      |     #log_info("gripper config:",to_str(GRIPPER_CONFIG_MAP[i]))
      |     if (GRIPPER_CONFIG_MAP[i].object == objectname):
      |         log_info("found gripper parameters [" + to_str(GRIPPER_CONFIG_MAP[i]) + "]")
      |         return GRIPPER_CONFIG_MAP[i]
      |     end
      |     i = i + 1
      | end
      | 
      | log_warning("no gripper parameters found for object type: " + to_str(objectname))
      | return create_gripper_config()
      | end
      | # Function to find a landmark by item
      | def find_landmark_by_id(lm_id):
      |     local i = 0
      |     while i < LANDMARK_MAP.length():
      |         if LANDMARK_MAP[i].lm_id == lm_id:
      |             log_info("found landmark with id(" + to_str(lm_id) + "): [" + to_str(LANDMARK_MAP[i].description) + "]")
      |             return LANDMARK_MAP[i]
      |         end
      |         i = i + 1
      |     end
      |     log_warning("landmark not found for lm_id [" + to_str(lm_id) + "]")
      |     return create_landmark()
      | end
      | # Function to find a landmark by item
      | def find_landmark_by_capture_pos(capture_pos):
      |     local i = 0
      |     while i < LANDMARK_MAP.length():
      |         if LANDMARK_MAP[i].capture_pos == capture_pos:
      |             log_info("found landmark by capture_pos [" + to_str(LANDMARK_MAP[i].description) + "]")
      |             return LANDMARK_MAP[i]
      |         end
      |         i = i + 1
      |     end
      |     log_warning("Landmark not found for capture_pos: [" + to_str(capture_pos) + "]")
      |     return create_landmark()
      | end
      | 
      | def update_landmark_by_capture_pos(capture_pos, lm_pos):
      |     local i = 0
      |     while i < LANDMARK_MAP.length():
      |         if LANDMARK_MAP[i].capture_pos == capture_pos:
      |             log_info("updated landmark from [" + to_str(LANDMARK_MAP[i].description) + "]")
      |             LANDMARK_MAP[i].actual_frame = lm_pos
      |             return True
      |         end
      |         i = i + 1
      |     end
      |     log_warning("Landmark not found for capture_pos: [" + to_str(capture_pos) + "]")
      |     return False
      | end
      | 
      | def update_landmark_by_id(lm_id,lm_pos):
      |     local i = 0
      |     while i < LANDMARK_MAP.length():
      |         if LANDMARK_MAP[i].lm_id == lm_id:
      |             log_info("updated landmark.actual_frame from [" + to_str(LANDMARK_MAP[i].description + "]"))
      |             LANDMARK_MAP[i].actual_frame = lm_pos
      |             return True
      |         end
      |         i = i + 1
      |     end
      |     log_warning("Landmark not found for lm_id " + to_str(lm_id))
      |     return False
      | end
      | 
      | def find_vision_config_by_frame(frame):
      |     local i = 0
      |     while i < VISION_CONFIG_MAP.length():
      |         if VISION_CONFIG_MAP[i].capture_pos == frame:
      |             log_info("Vision Config found: [" + to_str(VISION_CONFIG_MAP[i].description) + "]")
      |             return VISION_CONFIG_MAP[i]
      |         end
      |         i = i + 1
      |     end
      |     log_info("Vision Config not found for frame: " + to_str(frame))
      |     return create_vision_config()
      | end
      | 
      | def find_vision_config_by_itemid(id):
      |     local i = 0
      |     while i < VISION_CONFIG_MAP.length():
      |         if VISION_CONFIG_MAP[i].item_id == id:
      |             log_info("Vision Config found: [" + to_str(VISION_CONFIG_MAP[i].description) + "]")
      |             return VISION_CONFIG_MAP[i]
      |         end
      |         i = i + 1
      |     end
      |     log_info("Vision Config not found for item: " + to_str(id))
      |     return create_vision_config()
      | end
      | 
      | def find_inspect_config_by_itemid(id):
      |     local i = 0
      |     while i < INSPECT_CONFIG_MAP.length():
      |         if INSPECT_CONFIG_MAP[i].item_id == id:
      |             log_info("Inspect Config found: [" + to_str(INSPECT_CONFIG_MAP[i].description) + "]")
      |             return INSPECT_CONFIG_MAP[i]
      |         end
      |         i = i + 1
      |     end
      |     log_info("Inspect Config not found for item: " + to_str(id))
      |     return create_inspect_config()
      | end
    Script file /programs/04 Scripts/SCRIPT Device Robotiq Greifer v0.2.script
      | # ############ SCRIPT Device Robotiq Greifer ###############
      | # **********************************************************
      | # Customer          :   URG
      | # Product Name      :   uLabMobile
      | # **********************************************************
      | # Controller/Robot  :   UR5e
      | # Software          :   5.17
      | # Dependencies      :   Logs Script, Robotiq Gripper and Gripper Datastructure for args (Factory Script), URCAP Robotiq
      | # **********************************************************
      | # Author            :   D.Kreugel, P.Köhnke
      | # Copyright (c)     :   United Robotics Group Health and Food GmbH
      | #                       An der Riede 2
      | #                       28816 Stuhr
      | #                       Germany
      | # *********************************************************
      | # Description       :   Gripper Robotiq Device Interface for Robotiq E-Hand Gripper
      | # Version           :   0.2
      | # Created           :   18.07.2024
      | # Updated           :
      | # *********************************************************
      | # Modifications     :
      | #
      | # Date              :
      | # Name              :
      | # Reason            :
      | # *********************************************************
      | # TODO              :   documentation
      | 
      | # RobotiQ Gripper
      | ROBOTIQ_GRP_CLOSE = 0
      | ROBOTIQ_GRP_OPEN = 40
      | 
      | # #############FORCEMODE###############
      | ROBOTIQ_GRP_FORCE = struct(FULL=100, HALF=50, LOW=25, NONE=0)
      | 
      | # #############SPEED###################
      | ROBOTIQ_GRP_SPEED = struct(FAST=100, MEDIUM=50, SLOW=20)
      | 
      | # ############VALIDATION###############
      | ROBOTIQ_GRP_VALIDATION = struct(ON=1, OFF=0, SKIP=-1)
      | 
      | # struct(prepick=0, pick=0, place=0, force=0, speed=0, validation=0, object_type=0, description="default")
      | def gripper_robotiq_activate():
      |     return rq_activate_and_wait()
      | end
      | 
      | def gripper_robotiq_reset_and_activate():
      |     return rq_reset_and_activate()
      |     #return rq_reset()
      | end
      | 
      | def gripper_robotiq_is_activated():
      |     return rq_is_gripper_activated()
      | end
      | 
      | def gripper_robotiq_get_current_pos_mm():
      |     return rq_current_pos_mm()
      | end
      | # Function to check if the RobotiQ gripper has an object
      | def gripper_robotiq_has_object():
      |     result = rq_is_object_detected()
      |     if result == False:
      |         log_error("No object detected by the gripper")
      |     end
      |     return result
      | end
      | 
      | def gripper_robotiq_move_to_mm(mm):
      |     if(gripper_robotiq_is_activated() == False):
      |         gripper_robotiq_activate()
      |     end
      |     return rq_move_and_wait_mm(mm)
      | end
      | 
      | def gripper_robotiq_close():
      |     if(gripper_robotiq_is_activated() == False):
      |         gripper_robotiq_activate()
      |     end
      |     return rq_close_and_wait()
      | end
      | 
      | def gripper_robotiq_open():
      |     if(gripper_robotiq_is_activated() == False):
      |         gripper_robotiq_activate()
      |     end
      |     return rq_open_and_wait()
      | end
      | 
      | def gripper_robotiq_set_force(force):
      |     return rq_set_force_norm(force)
      | end
      | 
      | def gripper_robotiq_set_speed(velocity):
      |     return rq_set_speed_norm(velocity)
      | end
      | # Function to initialize the RobotiQ gripper
      | # args = struct(obj_type = object.obj_type, force = force, speed = speed, validation = validation, width = (prepick=2, pick=0, place=2))
      | def gripper_robotiq_init(args):
      |     log_info("args:"+to_str(args))
      |     gripper_robotiq_set_force(args.force)
      |     gripper_robotiq_set_speed(args.speed)
      |     if(gripper_robotiq_is_activated() == False):
      |         gripper_robotiq_activate()
      |     end
      |     log_info("Robotiq Gripper Initialized with arguments:" + to_str(args))
      |     return True
      | end
      | # Function to prepare the RobotiQ gripper for picking
      | # args = struct(obj_type = object.obj_type, force = force, speed = speed, validation = validation, width = (prepick=2, pick=0, place=2))
      | def gripper_robotiq_prepick(args):
      |     gripper_robotiq_init(args)
      | 
      |     if(args.width.prepick <= ROBOTIQ_GRP_CLOSE):
      |         rq_close_and_wait()
      |     elif(args.width.prepick >= ROBOTIQ_GRP_OPEN):
      |         rq_open_and_wait()
      |     else:
      |         rq_move_and_wait_mm(args.width.prepick)
      |     end
      | 
      |     log_info("Robotiq Gripper prepick with arguments:" + to_str(args))
      |     return True
      | end
      | 
      | # Function to place an object using the RobotiQ gripper
      | # args = struct(obj_type = object.obj_type, force = force, speed = speed, validation = validation, width = (prepick=2, pick=0, place=2))
      | def gripper_robotiq_place(args):
      |     gripper_robotiq_init(args)
      | 
      |     if(args.width.place <= ROBOTIQ_GRP_CLOSE):
      |         rq_close_and_wait()
      |     elif(args.width.place >= ROBOTIQ_GRP_OPEN):
      |         rq_open_and_wait()
      |     else:
      |         rq_move_and_wait_mm(args.width.place)
      |     end
      | 
      |     log_info("Gripper Place with arguments:"+ to_str(args))
      |     return True
      | end
      | 
      | # Function to pick an object using the RobotiQ gripper
      | # args = struct(obj_type = object.obj_type, force = force, speed = speed, validation = validation, width = (prepick=2, pick=0, place=2))
      | def gripper_robotiq_pick(args):
      |     gripper_robotiq_init(args)
      | 
      |     if(args.width.pick <= ROBOTIQ_GRP_CLOSE):
      |         rq_close_and_wait()
      |     elif(args.width.pick >= ROBOTIQ_GRP_OPEN):
      |         rq_open_and_wait()
      |     else:
      |         rq_move_and_wait_mm(args.width.pick)
      |     end
      | 
      |     log_info("Gripper Pick with arguments:" + to_str(args))
      | 
      |     if args.validation == ROBOTIQ_GRP_VALIDATION.ON:
      |         if gripper_robotiq_has_object() == False:
      |             log_error("Validation failed, no object detected")
      |             return False
      |         end
      |     end
      | 
      |     return True
      | end
      | 
      | 
      | # def gripper_robotiq_close_and_validate():
      | #     rq_close_and_wait()
      | #     if gripper_robotiq_has_object() == False:
      | #         log_error("Validation failed, no object detected")
      | #         return False
      | #     else:
      | #         return True
      | #     end
      | # end
    Script file /programs/04 Scripts/SCRIPT uLM Gripperconfig v0.6.script
      | ############# SCRIPT uLM Gripperconfig ###############
      | #*****************************************************
      | # Customer          :   URG
      | # Product Name      :   uLabMobile
      | #****************************************************
      | # Controller/Robot  :   UR5e
      | # Software          :   UR-Script
      | # Dependencies      :   physical Gripper and Datastructure from Factory for args -> Device Script and Implementations of the Functions
      | # How To            :   Assign all Functioncalls to the equivalent of the used Device Script
      | #****************************************************
      | # Author            :   D.Kreugel, P.Köhnke
      | # Copyright (c)     :   United Robotics Group Health and Food GmbH
      | #                       An der Riede 2
      | #                       28816 Stuhr
      | #                       Germany
      | #****************************************************
      | # Description       :   Defines all Gripperm related Parameters and Functions
      | # Version           :   0.6
      | # Created           :   18.07.2024
      | # Updated           :
      | #****************************************************
      | # Modifications     :   -> at the moment Gripperconfig linked to Robotiq Gripper Device Script
      | # Date              :   18.07.2017
      | # Name              :   D.Kreugel
      | # Reason            :   uLM Standard
      | #****************************************************
      | # TO DO             : Implement Activate and Reset Routine at the beginning or after an error depending on the state if an Object is gripped or not, documentation
      | 
      | 
      | 
      | # GRIPPER DEFINES
      | GRIPPER_CLOSE = ROBOTIQ_GRP_CLOSE
      | GRIPPER_OPEN = ROBOTIQ_GRP_OPEN
      | # #############FORCE###############
      | GRIPPER_FORCE = ROBOTIQ_GRP_FORCE
      | # #############SPEED###################
      | GRIPPER_SPEED = ROBOTIQ_GRP_SPEED
      | # ############VALIDATION###############
      | GRIPPER_VALIDATION = ROBOTIQ_GRP_VALIDATION
      | 
      | # takes force in %
      | def gripper_set_force(force):
      |     return gripper_robotiq_set_force(force)
      | end
      | 
      | # takes speed in %
      | def gripper_set_speed(velocity):
      |     return gripper_robotiq_set_speed(velocity)
      | end
      | 
      | def gripper_activate():
      |     return gripper_robotiq_activate()
      | end
      | 
      | def gripper_reset_and_activate():
      |     return gripper_robotiq_reset_and_activate()
      | end
      | 
      | def gripper_is_activated():
      |     return gripper_robotiq_is_activated()
      | end
      | 
      | def gripper_get_current_pos_mm():
      |     return gripper_robotiq_get_current_pos_mm()
      | end
      | 
      | def gripper_has_object():
      |     return gripper_robotiq_has_object()
      | end
      | 
      | def gripper_open():
      |     return gripper_robotiq_open()
      | end
      | 
      | def gripper_close():
      |     return gripper_robotiq_close()
      | end
      | 
      | def gripper_move_to_pos_mm(mm):
      |     return gripper_robotiq_move_to_mm(mm)
      | end
      | 
      | # args = struct(obj_type = object.obj_type, force = force, speed = speed, validation = validation, width = (prepick=2, pick=0, place=2))
      | def gripper_init(args):
      |     return gripper_robotiq_init(args)
      | end
      | 
      | # args = struct(obj_type = object.obj_type, force = force, speed = speed, validation = validation, width = (prepick=2, pick=0, place=2))
      | def gripper_prepick(args):
      |     return gripper_robotiq_prepick(args)
      | end
      | 
      | # args = struct(obj_type = object.obj_type, force = force, speed = speed, validation = validation, width = (prepick=2, pick=0, place=2))
      | def gripper_pick(args):
      |     return gripper_robotiq_pick(args)
      | end
      | 
      | # args = struct(obj_type = object.obj_type, force = force, speed = speed, validation = validation, width = (prepick=2, pick=0, place=2))
      | def gripper_place(args):
      |     return gripper_robotiq_place(args)
      | end
      | 
      | 
      | # def gripper_close_and_validate():
      | #     return gripper_robotiq_close_and_validate()
      | # end
    Script file /programs/04 Scripts/SCRIPT uLM Projectconfig 0.2.script
      | ############# SCRIPT uLM Projectconfig ###############
      | #*****************************************************
      | # Customer          :   URG
      | # Product Name      :   uLabMobile
      | #****************************************************
      | # Controller/Robot  :   UR5e
      | # Software          :   5.17
      | # Dependencies      :   Factory Script, Defines Script, relevant project knowledge about objects, patterns, items, commands, vision skills, landmarktypes and movements
      | # How To            :   Define Step by Step all Project Data by creating the objects and appending them to the assigned List, if you skip information
      | #                       the default value will be assigned -> give as many details as possible as the default values will not work in some cases
      | #****************************************************
      | # Author            :   D.Kreugel
      | # Copyright (c)     :   United Robotics Group Health and Food GmbH
      | #                       An der Riede 2
      | #                       28816 Stuhr
      | #                       Germany
      | #****************************************************
      | # Description       :   Project Related Configurations -> in the future will be configured by UGO
      | # Version           :   0.2
      | # Created           :   18.07.2024
      | # Updated           :
      | #****************************************************
      | # Modifications     :
      | # Date              :
      | # Name              :
      | # Reason            :
      | #****************************************************
      | # TO DO             :  Simplify Rack Assignment, create Enums for Choices that can be made and will be repeated in many projects, documentation
      | 
      | #
      | 
      | # Please Import DeviceScripts and Defines Script First as you may wanna use some of the Defined Variables here
      | 
      | # Define here the Objects that should be handled, add a new Object Type in the defines if necessary
      | # create_object(id=0, obj_name=0, height=0, width=0, color="default", material="default", description="default")
      | # struct(NONE=0, CC_SAMPLE=1, CC_RACK=2, COAG_SAMPLE=3, COAG_RACK=4, HEMA_SAMPLE=5, HEMA_RACK=6, INPUT_RACK=7, CF_RACK=8, ANY_SAMPLE=9, ANY_RACK=10)
      | #create_object(id=0, obj_name=0, height=0, width=0, obj_type = 0, description="default")
      | OBJECT_MAP.append(create_object(id=0, obj_name=Objects.NONE, obj_type=ObjectType.NONE, height=0, width=0, description="None Object"))
      | OBJECT_MAP.append(create_object(id=1, obj_name=Objects.CC_SAMPLE, obj_type=ObjectType.SAMPLE, height=108, width=15, description="BD Li-Heparin"))
      | OBJECT_MAP.append(create_object(id=2, obj_name=Objects.HEMA_SAMPLE, obj_type=ObjectType.SAMPLE, height=81, width=13, description="BD EDTA"))
      | OBJECT_MAP.append(create_object(id=3, obj_name=Objects.CC_SAMPLE, obj_type=ObjectType.SAMPLE, height=108, width=15, description="BD Li-Heparin"))
      | OBJECT_MAP.append(create_object(id=4, obj_name=Objects.HEMA_SAMPLE, obj_type=ObjectType.SAMPLE, height=81, width=13, description="Sarstedt EDTA"))
      | OBJECT_MAP.append(create_object(id=5, obj_name=Objects.CC_SAMPLE, obj_type=ObjectType.SAMPLE, height=110, width=15, description="Sarstedt Serum-Gel"))
      | OBJECT_MAP.append(create_object(id=6, obj_name=Objects.ANY_SAMPLE, obj_type=ObjectType.SAMPLE, height=110, width=15, description="Any Sample"))
      | OBJECT_MAP.append(create_object(id=7, obj_name=Objects.ANY_RACK, height=150, width=120, description="Any Rack"))
      | OBJECT_MAP.append(create_object(id=8, obj_name=Objects.CF_RACK, height=110, width=15, description="Centrifuge Rack"))
      | OBJECT_MAP.append(create_object(id=12, obj_name=Objects.COBAS_RACK, height=OBJECT_REFERENCE_HEIGHT, width=20, description="Cobas Rack"))
      | OBJECT_MAP.append(create_object(id=9, obj_name=Objects.TARA_SAMPLE, obj_type=ObjectType.SAMPLE, height=110, width=15, description="Tara Sample"))
      | OBJECT_MAP.append(create_object(id=10, obj_name=Objects.BUTTON, obj_type=ObjectType.BUTTON, height=0, width=0, description="Button"))
      | OBJECT_MAP.append(create_object(id=11, obj_name=Objects.XN550_DRAWER, height=OBJECT_REFERENCE_HEIGHT, width=25, description="XN550 Drawer"))
      | 
      | #create_sample(obj_id=0, diameter=0, color="", material="", description="")
      | SAMPLES = make_list(0,create_sample(),MAX_ITEM_OBJ)
      | SAMPLES.append(create_sample(obj_id=1, cap_diameter=17.4, raw_diameter=15.3, color="darkgreen", material="88", description="BD Li-Heparin -> decapped in Cobas"))
      | SAMPLES.append(create_sample(obj_id=1, cap_diameter=17.4, raw_diameter=15.3, color="darkgreen", material="80", description="BD Li-Heparin -> decapped in Cobas"))
      | SAMPLES.append(create_sample(obj_id=1, cap_diameter=17.4, raw_diameter=15.3, color="darkgreen", material="93", description="BD Li-Heparin -> decapped in archive"))
      | SAMPLES.append(create_sample(obj_id=2, cap_diameter=15.5, raw_diameter=12.3, color="violet", material="82", description="BD EDTA -> Sysmex ->Archive"))
      | SAMPLES.append(create_sample(obj_id=2, cap_diameter=15.5, raw_diameter=12.3, color="violet", material="91", description="BD EDTA ->Archive"))
      | SAMPLES.append(create_sample(obj_id=2, cap_diameter=15.5, raw_diameter=12.3, color="violet", material="96", description="BD EDTA ->Archive"))
      | SAMPLES.append(create_sample(obj_id=3, cap_diameter=17.4, raw_diameter=15.3, color="lightgreen", material="88", description="BD Li-Heparin -> decapped in Cobas"))
      | SAMPLES.append(create_sample(obj_id=3, cap_diameter=17.4, raw_diameter=15.3, color="lightgreen", material="93", description="BD Li-Heparin -> decapped in Archive"))
      | SAMPLES.append(create_sample(obj_id=3, cap_diameter=17.4, raw_diameter=15.3, color="lightgreen", material="97", description="BD Li-Heparin -> decapped in Archive"))
      | SAMPLES.append(create_sample(obj_id=4, cap_diameter=15.6, raw_diameter=12.3, color="red", material="82", description="BD EDTA -> Sysmex ->Archive"))
      | SAMPLES.append(create_sample(obj_id=4, cap_diameter=15.6, raw_diameter=12.3, color="red", material="91", description="BD EDTA -> Archive"))
      | SAMPLES.append(create_sample(obj_id=4, cap_diameter=15.6, raw_diameter=12.3, color="red", material="96", description="BD EDTA -> Archive"))
      | SAMPLES.append(create_sample(obj_id=5, cap_diameter=17.4, raw_diameter=15.3, color="brown", material="80", description="Sarstedt Serum-Gel -> decapped in Cobas"))
      | SAMPLES.append(create_sample(obj_id=5, cap_diameter=17.4, raw_diameter=15.3, color="brown", material="93", description="Sarstedt Serum-Gel -> decapped in Archive"))
      | 
      | # Gripper Configurations depending on the Object Type , add new force and speed in the Defines if necessary
      | # create_gripper_config(gripper_offset=struct(prepick=2, pick=0, place=2), force=0, speed=0, validation=0, object=create_object())
      | GRIPPER_CONFIG_MAP.append(create_gripper_config(gripper_offset=struct(prepick=2, pick=0, place=2), force=GRIPPER_FORCE.HALF, speed=GRIPPER_SPEED.MEDIUM, validation=GRIPPER_VALIDATION.ON, object=find_object_by_objectname(Objects.ANY_SAMPLE)))
      | GRIPPER_CONFIG_MAP.append(create_gripper_config(gripper_offset=struct(prepick=2, pick=0, place=2), force=GRIPPER_FORCE.FULL, speed=GRIPPER_SPEED.MEDIUM, validation=GRIPPER_VALIDATION.ON, object=find_object_by_objectname(Objects.ANY_RACK)))
      | GRIPPER_CONFIG_MAP.append(create_gripper_config(gripper_offset=struct(prepick=2, pick=0, place=2), force=GRIPPER_FORCE.HALF, speed=GRIPPER_SPEED.MEDIUM, validation=GRIPPER_VALIDATION.ON, object=find_object_by_objectname(Objects.CC_SAMPLE)))
      | GRIPPER_CONFIG_MAP.append(create_gripper_config(gripper_offset=struct(prepick=3, pick=0, place=3), force=GRIPPER_FORCE.HALF, speed=GRIPPER_SPEED.MEDIUM, validation=GRIPPER_VALIDATION.ON, object=find_object_by_objectname(Objects.HEMA_SAMPLE)))
      | GRIPPER_CONFIG_MAP.append(create_gripper_config(gripper_offset=struct(prepick=4, pick=0, place=4), force=GRIPPER_FORCE.HALF, speed=GRIPPER_SPEED.MEDIUM, validation=GRIPPER_VALIDATION.OFF, object=find_object_by_objectname(Objects.TARA_SAMPLE)))
      | GRIPPER_CONFIG_MAP.append(create_gripper_config(gripper_offset=struct(prepick=2, pick=0, place=2), force=GRIPPER_FORCE.FULL, speed=GRIPPER_SPEED.MEDIUM, validation=GRIPPER_VALIDATION.ON, object=find_object_by_objectname(Objects.CF_RACK)))
      | GRIPPER_CONFIG_MAP.append(create_gripper_config(gripper_offset=struct(prepick=2, pick=0, place=2), force=GRIPPER_FORCE.FULL, speed=GRIPPER_SPEED.MEDIUM, validation=GRIPPER_VALIDATION.ON, object=find_object_by_objectname(Objects.COBAS_RACK)))
      | GRIPPER_CONFIG_MAP.append(create_gripper_config(gripper_offset=struct(prepick=0, pick=0, place=0), force=GRIPPER_FORCE.HALF, speed=GRIPPER_SPEED.MEDIUM, validation=GRIPPER_VALIDATION.OFF, object=find_object_by_objectname(Objects.NONE)))
      | GRIPPER_CONFIG_MAP.append(create_gripper_config(gripper_offset=struct(prepick=0, pick=0, place=0), force=GRIPPER_FORCE.HALF, speed=GRIPPER_SPEED.MEDIUM, validation=GRIPPER_VALIDATION.OFF, object=find_object_by_objectname(Objects.BUTTON)))
      | GRIPPER_CONFIG_MAP.append(create_gripper_config(gripper_offset=struct(prepick=5, pick=25, place=5), force=GRIPPER_FORCE.HALF, speed=GRIPPER_SPEED.MEDIUM, validation=GRIPPER_VALIDATION.OFF, object=find_object_by_objectname(Objects.XN550_DRAWER)))
      | # create Patterns like Racks or Magazines
      | # easy if you define x and y regarding to the base coordinate system  if not you have to deal with transpose and or invert
      | # create_pattern(id=0, pattern_width=[0, 0], pattern_size=[0, 0], blocked=[-1, -1], obj_name=0, direction="X", transpose=False, invert=False, description="default")
      | # Objectss: NONE=0, CC_SAMPLE=1, CC_RACK=2, COAG_SAMPLE=3, COAG_RACK=4, HEMA_SAMPLE=5, HEMA_RACK=6, INPUT_RACK=7, CENTRIFUGE_RACK=8, ANY_SAMPLE=9, ANY_RACK=10
      | # ITEM_MODEL_MAP.append(create_pattern(id=0, pattern_width=[0, 0], pattern_size=[0, 0], blocked=[-1, -1, -1],  direction="X", transpose=False, invert=False, description="default"))
      | # ITEM_MODEL_MAP.append(create_pattern(id=1, pattern_width=[0.06, 0], pattern_size=[3, 1],  direction="X", description="Tara"))
      | # ITEM_MODEL_MAP.append(create_pattern(id=2, pattern_width=[0.183, 0.082], pattern_size=[10, 5], description="Sarstedt 50 D17 Rack"))
      | # ITEM_MODEL_MAP.append(create_pattern(id=3, pattern_width=[0.153, 0.067], pattern_size=[10, 5], description="Sarstedt 50 D13 Rack"))
      | # ITEM_MODEL_MAP.append(create_pattern(id=4, pattern_width=[0.06, 0.06], pattern_size=[3, 3], blocked=[5, -1, -1], description="Hettich Centrifuge Rack"))
      | # ITEM_MODEL_MAP.append(create_pattern(id=5, pattern_width=[0.093, 0.093], pattern_size=[2, 2],  description="Hettich Centrifuge Rack Magazin"))
      | # ITEM_MODEL_MAP.append(create_pattern(id=6, pattern_width=[0.08, 0.05], pattern_size=[5, 2], description="Sysmex XN 550 Rack"))
      | # ITEM_MODEL_MAP.append(create_pattern(id=7, pattern_width=[0.175, 0.078], pattern_size=[8, 4], description="URG Rack 40 D17"))
      | # ITEM_MODEL_MAP.append(create_pattern(id=8, pattern_width=[0.092, 0], pattern_size=[5, 1], description="Cobas Rack"))
      | # ITEM_MODEL_MAP.append(create_pattern(id=9, pattern_width=[0.245, 0.123], pattern_size=[3, 5], blocked=[9,11,12], description="Cobas Rack Magazin"))
      | # ITEM_MODEL_MAP.append(create_pattern(id=10, pattern_width=[0.237, 0.095], pattern_size=[11, 5], description="Atellica Rack 5x11"))
      | # ITEM_MODEL_MAP.append(create_pattern(id=11, pattern_width=[0.237, 0.095], pattern_size=[2, 2], description="Sensors LM"))
      | # ITEM_MODEL_MAP.append(create_pattern(id=12, pattern_width=[0.18, 0], pattern_size=[10, 1], description="Sysmex CS2500 Rack"))
      | # ITEM_MODEL_MAP.append(create_pattern(id=13, pattern_width=[0.310, 0.075], pattern_size=[13, 4], description="URG RACK 52 - Special Input"))
      | # ITEM_MODEL_MAP.append(create_pattern(id=14, pattern_width=[0.075, 0.075], pattern_size=[4, 6], description="URG RACK 24 - Special NoK"))
      | # ITEM_MODEL_MAP.append(create_pattern(id=15, pattern_width=[0.120, 0], pattern_size=[2, 1], description="XN550 Drawer"))
      | 
      | ITEM_MODEL_MAP.append(create_pattern(id=0, name="NONE", pattern_width=[0, 0], pattern_size=[0, 0], blocked=[-1, -1, -1],  direction="X", transpose=False, invert=False, description="default"))
      | ITEM_MODEL_MAP.append(create_pattern(id=1, name="TARA", pattern_width=[0.06, 0], pattern_size=[3, 1],  direction="X", description="Tara"))
      | ITEM_MODEL_MAP.append(create_pattern(id=4, name="CENTRIFUGE", pattern_width=[0.06, 0.06], pattern_size=[3, 3], blocked=[5, -1, -1], description="Hettich Centrifuge Rack"))
      | ITEM_MODEL_MAP.append(create_pattern(id=5, name="CENTRIFUGE_MAGAZINE", pattern_width=[0.093, 0.093], pattern_size=[2, 2],  description="Hettich Centrifuge Rack Magazin"))
      | ITEM_MODEL_MAP.append(create_pattern(id=6, name="SYSMEX_XN550", pattern_width=[0.08, 0.05], pattern_size=[5, 2], description="Sysmex XN 550 Rack"))
      | ITEM_MODEL_MAP.append(create_pattern(id=8, name="COBAS", pattern_width=[0.092, 0], pattern_size=[5, 1], description="Cobas Rack"))
      | ITEM_MODEL_MAP.append(create_pattern(id=9, name="COBAS_MAGAZINE", pattern_width=[0.245, 0.123], pattern_size=[3, 5], blocked=[9,11,12], description="Cobas Rack Magazin"))
      | ITEM_MODEL_MAP.append(create_pattern(id=13, name="INPUT", pattern_width=[0.310, 0.075], pattern_size=[13, 4], description="URG RACK 52 - Special Input"))
      | ITEM_MODEL_MAP.append(create_pattern(id=14, name="NOK", pattern_width=[0.075, 0.075], pattern_size=[4, 6], description="URG RACK 24 - Special NoK"))
      | ITEM_MODEL_MAP.append(create_pattern(id=15, name="DRAWER_XN550", pattern_width=[0.120, 0], pattern_size=[2, 1], description="XN550 Drawer"))
      | ITEM_MODEL_MAP.append(create_pattern(id=7, name="ARCHIVE", pattern_width=[0.175, 0.078], pattern_size=[8, 4], description="URG Rack 40 D17"))
      | 
      | 
      | 
      | 
      | 
      | 
      | # add a "skill" to the robots skillset the control system will send a string with the ls_item and action and here we will look if we have a matching skill to execute
      | # the item_modell defines the patterns which have to be used by the robot on multiple racks and or multiple samples in a rackpattern
      | # inner pattern is always dependung on the object that has to be moved and the outer pattern is the pattern for the containers where the objects are stored in.
      | # if racks have to be handled it is also an inner pattern cause the object to handle is the rack itself
      | # create_item(id=0, ls_item="default", frame=p[0,0,0,0,0,0], actionlist=create_action_list([]), item_model=create_item_model(), lm_id=0, description="default")
      | # create_item_model(inner=create_pattern(), outer=create_pattern(), description="default")
      | # ITEM_MAP.append(create_item(id=1, ls_item="Home", frame=F1_uLM_Home, actionlist=[ActionManipulator.MOVE_TO], description="uLM Move To Home"))
      | # ITEM_MAP.append(create_item(id=2, ls_item="InputStation", frame=F2_uLM_Input, actionlist=[ActionManipulator.PICK, ActionManipulator.PLACE], item_model=create_item_model(inner=Patterns.INPUT), description="uLM Pick and Place samples from Input"))
      | # ITEM_MAP.append(create_item(id=3, ls_item="InputCapture", frame=F3_Cap_Input, actionlist=[ActionCamera.INSPECT, ActionManipulator.MOVE_TO], description="uLM Inspect samples from Input and Move To Capture Position"))
      | # ITEM_MAP.append(create_item(id=4, ls_item="Bin", frame=F4_uLM_Bin, actionlist=[ActionManipulator.PLACE], description="uLM Place Cap to Bin"))
      | # ITEM_MAP.append(create_item(id=5, ls_item="StationaryGripper", frame=F5_uLM_Gripper, actionlist=[ActionManipulator.PICK, ActionManipulator.PLACE, ActionManipulator.DECAP, ActionManipulator.MOVE_TO, ActionManipulator.GRASP, ActionManipulator.RELEASE], description=" uLM stationary gripper"))
      | # ITEM_MAP.append(create_item(id=6, ls_item="CobasRack", frame=F6_uLM_Cobas_R, actionlist=[ActionManipulator.PICK, ActionManipulator.PLACE], item_model=create_item_model(outer=Patterns.COBAS_MAGAZINE), description="uLM Cobas Racks Pick and Place"))
      | # ITEM_MAP.append(create_item(id=7, ls_item="CobasMagazine", frame=F7_uLM_Coba_Mag, actionlist=[ActionManipulator.PICK, ActionManipulator.PLACE], item_model=create_item_model(inner=Patterns.COBAS, outer=Patterns.COBAS_MAGAZINE), description="uLM Cobas Magazine Samples Pick and Place"))
      | # ITEM_MAP.append(create_item(id=8, ls_item="DetectCobasRacks", frame=F8_Cap_Cobas_LM, actionlist=[ActionCamera.DETECT_OBJECTS, ActionManipulator.MOVE_TO], lm_id=2, description="uLM Cobas Rack Detection and Move To Capture"))
      | # ITEM_MAP.append(create_item(id=9, ls_item="TaraMagazine", frame=F9_uLM_Tara, actionlist=[ActionManipulator.PICK, ActionManipulator.PLACE], item_model=create_item_model(inner=Patterns.TARA), description="uLM Centrifuge Tara Pick and Place"))
      | # ITEM_MAP.append(create_item(id=10, ls_item="CentrifugeCapture", frame=F10_Cap_CF, actionlist=[ActionManipulator.MOVE_TO, ActionCamera.DETECT], lm_id=1, description="Centrifuge Device Move to Capture Pos and Detect Landmarks"))
      | # ITEM_MAP.append(create_item(id=11, ls_item="Centrifuge", frame=F11_CF_PiPl, actionlist=[ActionManipulator.PICK, ActionManipulator.PLACE], description="Centrifuge Device Rack Pick and Place"))
      | # ITEM_MAP.append(create_item(id=12, ls_item="CentrifugeMagazine", frame=F12_uLM_CF_Mag, actionlist=[ActionManipulator.PICK, ActionManipulator.PLACE], item_model=create_item_model(inner=Patterns.CENTRIFUGE, outer=Patterns.CENTRIFUGE_MAGAZINE), description=" uLM Centrifuge Magazin Pick and Place"))
      | # ITEM_MAP.append(create_item(id=13, ls_item="CentrifugeRack", frame=F13_uLM_CF_R, actionlist=[ActionManipulator.PICK, ActionManipulator.PLACE], item_model=create_item_model(outer=Patterns.CENTRIFUGE_MAGAZINE), description="uLM Centrifuge Magazin Pick and Place Racks"))
      | # ITEM_MAP.append(create_item(id=14, ls_item="DailyArchive", frame=F14_uLM_Archive, actionlist=[ActionManipulator.PICK, ActionManipulator.PLACE], item_model=create_item_model(inner=Patterns.ARCHIVE), description="uLM Pick and Place samples from Archive Rack"))
      | # ITEM_MAP.append(create_item(id=15, ls_item="NokRack", frame=F15_uLM_Nok, actionlist=[ActionManipulator.PICK, ActionManipulator.PLACE], item_model=create_item_model(inner=Patterns.NOK), description="uLM Pick and Place samples from Nok Rack"))
      | # ITEM_MAP.append(create_item(id=16, ls_item="CobasInput", frame=F16_Cobas_Input, actionlist=[ActionManipulator.PLACE], description="uLM Place Cobasrack in Cobas Device"))
      | # ITEM_MAP.append(create_item(id=17, ls_item="CobasInputCapture", frame=F17_Cobas_Cap, actionlist=[ActionCamera.DETECT, ActionManipulator.MOVE_TO], lm_id=3, description="uLM Place Cobasrack in Cobas Device"))
      | # ITEM_MAP.append(create_item(id=18, ls_item="XN550Input", frame=F18_XN550_Input, actionlist=[ActionManipulator.PICK, ActionManipulator.PLACE], item_model=create_item_model(inner=Patterns.SYSMEX_XN550, outer=Patterns.DRAWER_XN550), lm_id=4, description="uLM Pick and Place Samples in or out of XN550 Racks"))
      | # ITEM_MAP.append(create_item(id=19, ls_item="XN550Capture", frame=F19_XN550_Cap, actionlist=[ActionCamera.DETECT, ActionManipulator.MOVE_TO], lm_id=4, description="uLM Move To and Capture LM XN550"))
      | # ITEM_MAP.append(create_item(id=20, ls_item="XN550Drawer", frame=F20_XN550_Draw, actionlist=[ActionManipulator.DRAWER_OPEN, ActionManipulator.DRAWER_CLOSE], item_model=create_item_model(inner=Patterns.DRAWER_XN550), lm_id=4, description="uLM Open and close Drawer XN550"))
      | # ITEM_MAP.append(create_item(id=21, ls_item="XN550Button", frame=F21_XN550_Btn, actionlist=[ActionManipulator.PUSH], lm_id=4, description="uLM Push XN550 Button"))
      | # ITEM_MAP.append(create_item(id=22, ls_item="AMR", frame=p[0,0,0,0,0,0], actionlist=[ActionAMR.READ, ActionAMR.LOAD_MISSION, ActionAMR.START_MISSION, ActionAMR.NAVIGATE, ActionAMR.ACKNOWLEDGE], description="all AMR actions"))
      | 
      | 
      | 
      | # ITEM_MAP.append(create_item(id=31, ls_item="TestLM", frame=TestLM, actionlist=[ActionManipulator.PICK, ActionManipulator.PLACE], item_model=create_item_model(inner=Rack.SYSMEX_CS2500), lm_id=5, description="LM Test"))
      | # Fills the Vision Config List with Projectrelated Data
      | # workspaceid and skillid are highly robominds related so probably will not stay like this in the future
      | # sample detection: dx and dy are used to calculate the positions in a rack and given by the offset which will be applied in order to assign the sample to a place in the rack
      | # create_vision_config(workspace_id="", skill_id="", item_id=-1, capture_pos=p[0,0,0,0,0,0], dx=0, dy=0, target_origin=p[0,0,0,0,0,0], selector="default", description="default")
      | # VISION_CONFIG_MAP.append(create_vision_config(workspace_id="96017791-f581-4e9e-93da-6951695fccc8", skill_id="8885cfe1-6784-4293-bd26-52ebdc67bf95", capture_pos=F10_Cap_CF, target_origin=p[0,0,0,0,0,0], item_id=11, description="LM Detect CF"))
      | # VISION_CONFIG_MAP.append(create_vision_config(workspace_id="96017791-f581-4e9e-93da-6951695fccc8", skill_id="8885cfe1-6784-4293-bd26-52ebdc67bf95", capture_pos=F8_Cap_Cobas_LM, target_origin=p[0,0,0,0,0,0], item_id=8, description="LM Detect Cobas Racks"))
      | # VISION_CONFIG_MAP.append(create_vision_config(workspace_id="8f0ad01c-dc36-4fdd-b295-0b6b4a38b89a", skill_id="afdc9e13-ea83-40d6-a805-bb041453d2e5", capture_pos=F3_Cap_Input, target_origin=F2_uLM_Input, item_id=3, description="Lab Solution Input Capture"))
      | # VISION_CONFIG_MAP.append(create_vision_config(workspace_id="96017791-f581-4e9e-93da-6951695fccc8", skill_id="8885cfe1-6784-4293-bd26-52ebdc67bf95", capture_pos=F19_XN550_Cap, target_origin=F18_XN550_Input, item_id=18, description="Input XN550"))
      | # VISION_CONFIG_MAP.append(create_vision_config(workspace_id="96017791-f581-4e9e-93da-6951695fccc8", skill_id="8885cfe1-6784-4293-bd26-52ebdc67bf95", capture_pos=F19_XN550_Cap, target_origin=POS_Z, item_id=19, description="LM Detect XN550F"))
      | # VISION_CONFIG_MAP.append(create_vision_config(workspace_id="96017791-f581-4e9e-93da-6951695fccc8", skill_id="8885cfe1-6784-4293-bd26-52ebdc67bf95", capture_pos=F10_Cap_CF, target_origin=POS_Z, item_id=10, description="LM Detect CF"))
      | # VISION_CONFIG_MAP.append(create_vision_config(workspace_id="96017791-f581-4e9e-93da-6951695fccc8", skill_id="8885cfe1-6784-4293-bd26-52ebdc67bf95", capture_pos=F19_XN550_Cap, target_origin=F20_XN550_Draw, item_id=20, description="Drawer XN550"))
      | # VISION_CONFIG_MAP.append(create_vision_config(workspace_id="96017791-f581-4e9e-93da-6951695fccc8", skill_id="8885cfe1-6784-4293-bd26-52ebdc67bf95", capture_pos=F19_XN550_Cap, target_origin=F21_XN550_Btn, item_id=21, description="Button XN550"))
      | # VISION_CONFIG_MAP.append(create_vision_config(workspace_id="96017791-f581-4e9e-93da-6951695fccc8", skill_id="8885cfe1-6784-4293-bd26-52ebdc67bf95", capture_pos=TestLMCap, target_origin=p[0,0,0,0,0,0], item_id=30, description="Button XN550"))
      | # VISION_CONFIG_MAP.append(create_vision_config(workspace_id="96017791-f581-4e9e-93da-6951695fccc8", skill_id="8885cfe1-6784-4293-bd26-52ebdc67bf95", capture_pos=TestLMCap, target_origin=TestLM, item_id=31, description="Button XN550"))
      | 
      | # VISION_CONFIG_MAP.append(create_vision_config(workspace_id="96017791-f581-4e9e-93da-6951695fccc8", skill_id="8885cfe1-6784-4293-bd26-52ebdc67bf95", target_origin=p[0,0,0,0,0,0], item_id=11, description="LM Detect CF"))
      | # VISION_CONFIG_MAP.append(create_vision_config(workspace_id="96017791-f581-4e9e-93da-6951695fccc8", skill_id="8885cfe1-6784-4293-bd26-52ebdc67bf95", target_origin=p[0,0,0,0,0,0], item_id=8, description="LM Detect Cobas Racks"))
      | # VISION_CONFIG_MAP.append(create_vision_config(workspace_id="8f0ad01c-dc36-4fdd-b295-0b6b4a38b89a", skill_id="afdc9e13-ea83-40d6-a805-bb041453d2e5", target_origin=F2_uLM_Input, item_id=3, description="Lab Solution Input Capture"))
      | # VISION_CONFIG_MAP.append(create_vision_config(workspace_id="96017791-f581-4e9e-93da-6951695fccc8", skill_id="8885cfe1-6784-4293-bd26-52ebdc67bf95", target_origin=F18_XN550_Input, item_id=18, description="Input XN550"))
      | # VISION_CONFIG_MAP.append(create_vision_config(workspace_id="96017791-f581-4e9e-93da-6951695fccc8", skill_id="8885cfe1-6784-4293-bd26-52ebdc67bf95", target_origin=POS_Z, item_id=19, description="LM Detect XN550F"))
      | # VISION_CONFIG_MAP.append(create_vision_config(workspace_id="96017791-f581-4e9e-93da-6951695fccc8", skill_id="8885cfe1-6784-4293-bd26-52ebdc67bf95", target_origin=POS_Z, item_id=10, description="LM Detect CF"))
      | # VISION_CONFIG_MAP.append(create_vision_config(workspace_id="96017791-f581-4e9e-93da-6951695fccc8", skill_id="8885cfe1-6784-4293-bd26-52ebdc67bf95", target_origin=F20_XN550_Draw, item_id=20, description="Drawer XN550"))
      | # VISION_CONFIG_MAP.append(create_vision_config(workspace_id="96017791-f581-4e9e-93da-6951695fccc8", skill_id="8885cfe1-6784-4293-bd26-52ebdc67bf95", target_origin=F21_XN550_Btn, item_id=21, description="Button XN550"))
      | # VISION_CONFIG_MAP.append(create_vision_config(workspace_id="96017791-f581-4e9e-93da-6951695fccc8", skill_id="8885cfe1-6784-4293-bd26-52ebdc67bf95", target_origin=p[0,0,0,0,0,0], item_id=30, description="Button XN550"))
      | # VISION_CONFIG_MAP.append(create_vision_config(workspace_id="96017791-f581-4e9e-93da-6951695fccc8", skill_id="8885cfe1-6784-4293-bd26-52ebdc67bf95", target_origin=TestLM, item_id=31, description="Button XN550"))
      | 
      | # local inputrack = find_pattern_by_name("INPUT")
      | # INSPECT_CONFIG_MAP.append(create_inspect_config(item_id=3, dx=inputrack.pattern_width[0]/(inputrack.pattern_size[0]-1), dy=inputrack.pattern_width[1]/(inputrack.pattern_size[1]-1), rack_size=inputrack.pattern_size , description="Input Capture"))
      | # # Fills the Landmark List with Projectrelated Data
      | # # create_landmark(lm_id=0, marker_id=-1, marker_size=0.1, marker_type="aruco_7x7", capture_pos=p[0,0,0,0,0,0], init_frame=p[0,0,0,0,0,0], search_offset=[0,0,0], actual_frame=p[0,0,0,0,0,0], description="")
      | # LANDMARK_MAP.append(create_landmark(lm_id=1, marker_id=3, marker_size=0.1, marker_type="aruco_7x7", capture_pos = F10_Cap_CF, init_frame=p[-0.617789, -0.065471, 0.07918, 0.020983, -0.012695, 1.512066], search_offset=[0.15, 0.15, 0.1], actual_frame=p[-0.617789, -0.065471, 0.07918, 0.020983, -0.012695, 1.512066], description="LM CF Lid"))
      | # LANDMARK_MAP.append(create_landmark(lm_id=2, marker_id=-1, marker_size=0.0085, marker_type="aruco_4x4", capture_pos = F8_Cap_Cobas_LM, init_frame=p[0,0,0,0,0,0], search_offset=[0.15, 0.15, 0.1], actual_frame=POS_Z, description="LM Cobas Rack Detection"))
      | # LANDMARK_MAP.append(create_landmark(lm_id=3, marker_id=0, marker_size=0.1, marker_type="aruco_7x7", capture_pos = F17_Cobas_Cap, init_frame=p[-0.667,-0.194,0.100,0,0,0], search_offset=[0.15, 0.15, 0.1], actual_frame=POS_Z, description="LM Cobas Cap"))
      | # LANDMARK_MAP.append(create_landmark(lm_id=4, marker_id=4, marker_size=0.1, marker_type="aruco_7x7", capture_pos = F19_XN550_Cap, init_frame=p[0.124,-0.976,0.355,-0.008,0.025,3.131], search_offset=[0.15, 0.15, 0.1], actual_frame=p[0,0,0,0,0,0], description="LM XN550 Cap"))
      | # LANDMARK_MAP.append(create_landmark(lm_id=5, marker_id=0, marker_size=0.1, marker_type="aruco_7x7", capture_pos = TestLMCap, init_frame=p[-0.49,-0.144,0.092,0,-0.008,0.001], search_offset=[0.15, 0.15, 0.1], actual_frame=POS_Z, description="LM Test"))
      | # # Configuration of all movement related parameters
      | # # create_movement(id=0, hh_approach=POS_Z, h_approach=POS_Z, approach=POS_Z, h_target=POS_Z, target=POS_Z, retract=POS_Z, h_retract=POS_Z, hh_retract=POS_Z, h_frame=POS_Z, frame=POS_Z, speed=1, acceleration=1, description="default")
      | # MOVEMENT_MAP.append(create_movement(description="TestLMCap", frame=TestLMCap, actionlist=[ActionManipulator.MOVE_TO]))
      | # MOVEMENT_MAP.append(create_movement(description="TestLM", frame=TestLM, actionlist=[ActionManipulator.PICK,ActionManipulator.PLACE],
      | #         approach=p[0,0,0.1,0,0,0],
      | #         retract=p[0,0,0.1,0,0,0]))
      | # MOVEMENT_MAP.append(create_movement(description="Home - MOVE_TO", frame=F1_uLM_Home, actionlist=[ActionManipulator.MOVE_TO]))
      | # MOVEMENT_MAP.append(create_movement(description="Input - PICK&PLACE", frame=F2_uLM_Input, actionlist=[ActionManipulator.PICK,ActionManipulator.PLACE],
      | #         approach=p[0,0,0.1,0,0,0],
      | #         retract=p[0,0,0.1,0,0,0]))
      | # MOVEMENT_MAP.append(create_movement(description="Capture Input - MOVE_TO", frame=F3_Cap_Input, actionlist=[ActionManipulator.MOVE_TO]))
      | # MOVEMENT_MAP.append(create_movement(description="BIN - PLACE", frame=F4_uLM_Bin, actionlist=[ActionManipulator.PLACE],
      | #         approach=p[0,0,0.1,0,0,0],
      | #         retract=p[0,0,0.1,0,0,0]))
      | # MOVEMENT_MAP.append(create_movement(description="Gripper - Move To", frame=F5_uLM_Gripper, actionlist=[ActionManipulator.MOVE_TO],
      | #         approach=p[0,0,0.1,0,0,0]))
      | # MOVEMENT_MAP.append(create_movement(description="Gripper - Pick", frame=F5_uLM_Gripper, actionlist=[ActionManipulator.PICK],
      | #         retract=p[0,0,0.1,0,0,0]))
      | # MOVEMENT_MAP.append(create_movement(description="Gripper - Place", frame=F5_uLM_Gripper, actionlist=[ActionManipulator.PLACE],
      | #         approach=p[0,0,0.1,0,0,0]))
      | # MOVEMENT_MAP.append(create_movement(description="CobasRack Pick & Place", frame=F6_uLM_Cobas_R, actionlist=[ActionManipulator.PICK,ActionManipulator.PLACE],
      | #         approach=p[0,0,0.1,0,0,0],
      | #         target=p[0,0,0,0,0,d2r(90)],
      | #         retract=p[0,0,0.1,0,0,0]))
      | # MOVEMENT_MAP.append(create_movement(description="CobasMagazine Pick & Place", frame=F7_uLM_Coba_Mag, actionlist=[ActionManipulator.PICK,ActionManipulator.PLACE],
      | #         approach=p[0,0,0.1,0,0,0],
      | #         target=p[0,0,0,0,0,-d2r(90)],
      | #         retract=p[0,0,0.1,0,0,0]))
      | # MOVEMENT_MAP.append(create_movement(description="Capture Position Cobas Landmarks", frame=F8_Cap_Cobas_LM, actionlist=[ActionManipulator.MOVE_TO]))
      | # MOVEMENT_MAP.append(create_movement(description="TaraMagazine - PICK & PLACE", frame=F9_uLM_Tara, actionlist=[ActionManipulator.PICK,ActionManipulator.PLACE],
      | #         approach=p[0,0,0.13,0,0,0],
      | #         target=p[0,0,0,0,0,-d2r(90)],
      | #         retract=p[0,0,0.13,0,0,0]))
      | # MOVEMENT_MAP.append(create_movement(description="Capture Position - Centrifuge LM", frame=F10_Cap_CF,actionlist=[ActionManipulator.MOVE_TO]))
      | # MOVEMENT_MAP.append(create_movement(description="Pick and Place Racks - Centrifuge Lid", frame=F11_CF_PiPl, actionlist=[ActionManipulator.PICK,ActionManipulator.PLACE],
      | #         approach=p[0,0,0.3,0,0,0],
      | #         retract=p[0,0,0.3,0,0,0]))
      | # MOVEMENT_MAP.append(create_movement(description="Pick and Place Samples - Centrifuge on uLM", frame=F12_uLM_CF_Mag, actionlist=[ActionManipulator.PICK,ActionManipulator.PLACE],
      | #         approach=p[0,0,0.13,0,0,0],
      | #         retract=p[0,0,0.13,0,0,0]
      | #         ))
      | # MOVEMENT_MAP.append(create_movement(description="Pick and Place Racks - Centrifuge on uLM", frame=F13_uLM_CF_R, actionlist=[ActionManipulator.PICK,ActionManipulator.PLACE],
      | #         approach=p[0,0,0.15,0,0,0],
      | #         retract=p[0,0,0.15,0,0,0]
      | #         ))
      | 
      | # MOVEMENT_MAP.append(create_movement(description="Pick and Place Samples XN550 Racks in Device", frame=F18_XN550_Input, actionlist=[ActionManipulator.PICK,ActionManipulator.PLACE],
      | #         approach=p[0,0,0.1,0,0,0],
      | #         target = p[0,0,0,0,0,d2r(90)],
      | #         retract=p[0,0,0.1,0,0,0]
      | #         ))
      | # MOVEMENT_MAP.append(create_movement(description="Capture LM XN550", frame=F19_XN550_Cap, actionlist=[ActionManipulator.MOVE_TO]))
      | # MOVEMENT_MAP.append(create_movement(description="Open XN550 Drawer ", frame=F20_XN550_Draw, actionlist=[ActionManipulator.DRAWER_OPEN],
      | #         h_approach=p[0.07,0,0.1,0,0,0],
      | #         approach=p[0,0,0.1,0,0,0],
      | #         target = p[0,0,0,0,0,d2r(90)],
      | #         retract=p[0.07,0,0,0,0,0],
      | #         h_retract=p[0.07,0,0.1,0,0,0]
      | #         ))
      | # MOVEMENT_MAP.append(create_movement(description="Close XN550 Drawer ", frame=F20_XN550_Draw, actionlist=[ActionManipulator.DRAWER_CLOSE],
      | #         h_approach=p[0.07,0,0.1,0,0,0],
      | #         approach=p[0.07,0,0,0,0,0],
      | #         target = p[0,0,0,0,0,d2r(90)],
      | #         retract=p[0,0,0.1,0,0,0],
      | #         h_retract=p[0.07,0,0.1,0,0,0]
      | #         ))
      | # MOVEMENT_MAP.append(create_movement(description="Push XN550 Button ", frame=F21_XN550_Btn, actionlist=[ActionManipulator.PUSH],
      | #         approach=p[0,0,0.15,0,0,0],
      | #         retract=p[0,0,0.15,0,0,0]
      | #         ))
      | # MOVEMENT_MAP.append(create_movement(description="Capture Position 2 Input", frame=F_Cap_Input2,actionlist=[ActionManipulator.MOVE_TO]))
    Script file /programs/04 Scripts/SCRIPT Objects V0.1.script
      | #*****************************************************
      | # customer          :   INTERNAL
      | # project name      :
      | #****************************************************
      | # controller        :   UR
      | # software          :   5.17.3
      | #****************************************************
      | # author            :   P. Koehnke
      | # Copyright (c)     :   United Robotics Group
      | #                       An der Riede 2
      | #                       28816 Stuhr
      | #                       Germany
      | #****************************************************
      | # description       :   object database
      | # version:      	:   0.1
      | # created           :   09.10.2024
      | # updated           :
      | #****************************************************
      | # modifications     :
      | #
      | # date              :
      | # name              :
      | # reason            :
      | #****************************************************
      | 
      | def create_object_2(id=0, name="", type=0, dimension=struct(length=0, width=0, height=0, diameter=0), gripper_offset=p[0,0,0,0,0,0]):
      |     return struct(id=id, name=name, type=type, dimension=dimension, gripper_offset=gripper_offset)
      | end
      | 
      | OBJ = create_object_2()
      | OBJs = make_list(0, create_object_2(), 50)
      | 
      | OBJs.append(create_object_2(id=1, name="rack centrifuge", type=1, dimension=struct(length=0, width=0, height=0.106, diameter=0.020), gripper_offset=p[0,0,0.095,0,0,2.356]))
      | OBJs.append(create_object_2(id=2, name="sample tube 1", type=2, dimension=struct(length=0, width=0, height=0.106, diameter=0.015), gripper_offset=p[0,0,0,0,0,0]))
      | OBJs.append(create_object_2(id=3, name="rack sarstedt", type=3, dimension=struct(length=0, width=0, height=0.100, diameter=0.020), gripper_offset=p[0,0,0,0,0,0]))
      | def create_jig_2(id=0, name="", type=0, capacity=0, jig_offset=p[0,0,0,0,0,0]):
      |     # iformation about used jigs
      |     return struct(id=id, name=name, type=type, capacity=capacity, jig_offset=jig_offset)
      | end
      | 
      | JIG2 = create_jig_2()
      | JIGs = make_list(0, create_jig_2(), 10)
      | 
      | JIGs.append(create_jig_2(id=1, name="3FG", type=1, capacity=1, jig_offset=p[0,0,0,0,0,0]))
      | JIGs.append(create_jig_2(id=2, name="jig input", type=2, capacity=1, jig_offset=p[0,0,0,0,0,-3.927]))
      | JIGs.append(create_jig_2(id=3, name="jig output", type=3, capacity=1, jig_offset=p[0,0,0,0,0,0.78]))
      | JIGs.append(create_jig_2(id=4, name="jig centrifuge racks", type=4, capacity=4, jig_offset=p[0,0,0,0,0,-3.9162]))
      | JIGs.append(create_jig_2(id=6, name="jig bin", type=6, capacity=1, jig_offset=p[0,0,0,0,0,0]))
      | JIGs.append(create_jig_2(id=7, name="jig sarstedt racks", type=7, capacity=1, jig_offset=p[0,0,-0.02,0,0,0]))
  Folder BeforeStarts [hidden by the author, left out]
Robot Program (runOnlyOnce=false)
  Folder MAIN
    Script: command_manager(external_control="uGO", cond_suspend=(ITM_Manipulated and AMR_AtTarget and AMR_Charging and AMR_Battery<40), cond_unsuspend=(AMR_Battery≟60))
    Script: log_state(STATE_Info)
    Switch expression=STATE
      Case (caseValue=1)
        Folder Stopping
          STATE_Info := "Stopping"
          Script: end_freedrive_mode()
          Set NoAction tcp=TCP
          PSE_T := get_tool_free_pose(dir=[0,0,0.150], move_in_base_frame=True)
          If is_reachable(Base, [PSE_T])
            MoveL speed 150 mm/s, acceleration 1200 mm/s^2 (useActiveTCP=true) feature=Base
              Waypoint Variable (Variable): variable=PSE_T
          Script: do_transition(keep_rxry=OBJ_Picked, r=0)
          Folder Decapper [hidden by the author, left out]
          SuppressedNode
            Folder Centrifuge [hidden by the author, left out]
          Call Sub_AMR_MiR_V3
          If stopping() and AMR_Done
            STATE := 2
            Script: ugo_update_outputs()
      Case (caseValue=2)
        Folder Stopped
          STATE_Info := "Stopped"
          Call Sub_AMR_MiR_V3
          If CMD_Reset
            STATE := 3
            Script: ugo_update_outputs()
      Case (caseValue=3)
        Folder  Resetting [hidden by the author, left out]
      Case (caseValue=4)
        Folder Idle [hidden by the author, left out]
      Case (caseValue=5)
        Folder Starting
          STATE_Info := "Starting"
          'ADD COMMANDS WHAT TO START WITH'
          Call Sub_AMR_MiR_V3
          Folder get ugo data
            Folder Assign Tasks
              Script: TASK.ID = ugo_get_task()
              If TASK.ID≟1
                Task_info := "Charge"
                Folder Parameters
                  AMR_PosTarget := 1
              ElseIf TASK.ID≟9
                'Pick Sarstedt Rack from Variable source'
                Task_info := "Navigate to Target"
                Folder Parameters
                  AMR_PosTarget := UGO.read_input("00","ITM_ID")
              ElseIf TASK.ID≟10
                'Pick Sarstedt Rack from Variable source'
                Task_info := "Pick Rack"
                AMR_PosTarget := AMR_PosActual
                Folder Parameters
                  ITM_ID := UGO.read_input("00","ITM_ID")
                  JIG := UGO.read_input("00","JIG_ID")
                  OBJ_Type := 3
                SuppressedNode
                  ITM_ID := 1
              ElseIf TASK.ID≟11
                'Place Sarstedt Rack on Variable target'
                Task_info := "Place Rack"
                Folder Parameters
                  ITM_ID := UGO.read_input("00","ITM_ID")
                  JIG := UGO.read_input("00","JIG_ID")
                  OBJ_Type := 3
                SuppressedNode
                  ITM_ID := 1
              SuppressedNode
                ElseIf TASK.ID≟12
                  Task_info := "Decapping"
                  Folder Parameters
                    ITM_ID := 1
                    AMR_PosTarget := AMR_PosActual
                    SuppressedNode
                      PRC_TubCounter := 0
              ElseIf TASK.ID≟13
                Task_info := "Empty racks"
                Folder Parameters
                  ITM_ID := 1
                  AMR_PosTarget := AMR_PosActual
              ElseIf TASK.ID≟14
                Task_info := "Decap"
                Folder Parameters
                  ITM_ID := 1
                  OBJ_Type := 2
                  JIG := 7
                  AMR_PosTarget := AMR_PosActual
              ElseIf TASK.ID≟99
                Task_info := "Decapping and barcode alignment"
                Folder Parameters
                  PRC_TubNumber := UGO.read_input("00","TubesNb")
                  PRC_TubCounter := 0
                  ITM_ID := 1
                  AMR_PosTarget := AMR_PosActual
              SuppressedNode
                ElseIf TASK.ID≟14
                  Task_info := "Load Centrifuge"
                  Folder Parameters
                    PRC_RackCounter := 0
                    Script: TASK.WORK.ITM_ID_Src=1
                    Script: TASK.WORK.ITM_ID_Tgt=2
                    AMR_PosTarget := 4
                    AMR_FootprintID := 1
              ElseIf TASK.ID≟15
                Task_info := "Unoad Centrifuge"
                Folder Parameters
                  PRC_RackCounter := 0
                  Script: TASK.WORK.ITM_ID_Src=2
                  Script: TASK.WORK.ITM_ID_Tgt=1
                  AMR_PosTarget := 4
                  AMR_FootprintID := 1
              SuppressedNode
                ElseIf TASK.ID≟99
                  Task_info := "Load Biorad"
                  Folder Parameters
                    PRC_RackCounter := 0
                    ITM_ID := 2
                    CAM_LM_ID := 0
                    SuppressedNode
                      AMR_PosTarget := 1
                    AMR_PosTarget := AMR_PosActual
                    PRC_RackNumber := UGO.read_input("00","RackNb")
              SuppressedNode
                ElseIf TASK.ID≟99
                  Task_info := "Unload Biorad"
                  Folder Parameters
                    PRC_RackCounter := 0
                    ITM_ID := 2
                    CAM_LM_ID := 0
                    SuppressedNode
                      AMR_PosTarget := 1
                    AMR_PosTarget := AMR_PosActual
                    PRC_RackNumber := UGO.read_input("00","RackNb")
              Else 
                Script: set_error(ERROR_WRONG_ORDER)
          Folder test ugo
            Wait Sleep waitTime=0.2
            Script: ugo_update_outputs()
          If starting() and AMR_Done
            Script: log_message(Task_info, "New Task: ")
            Script: log_message(to_str(TASK.ID), "Task_ID: ")
            Script: do_transition(keep_rxry=OBJ_Picked)
            STATE := 6
            Script: ugo_update_outputs()
      Case (caseValue=6)
        Folder Execute
          STATE_Info := "Execute"
          If not CMD_Hold and not CMD_Suspend (checkContinuously=true)
            Switch expression=PROCESS_Step
              Case (caseValue=0)
                PROCESS_Info := "process control"
                Script: log_process(PROCESS_Info)
                Folder process control
                  If not AMR_AtTarget
                    PROCESS_Step := 1
                  ElseIf (( not ITM_Prepared and  not WRK_Done) or (ITM_Prepared and WRK_Done))
                    PROCESS_Step := 2
                  ElseIf not WRK_Done
                    PROCESS_Step := 3
                  Else 
                    Folder task finished
                      PROCESS_Info := ""
                      STATE := 7
                      Script: ugo_update_outputs()
              Case (caseValue=1)
                Folder navigate
                  'MOVING THE uML'
                  PROCESS_Info := "move to target"
                  Script: log_process(PROCESS_Info)
                  If TASK.ID≟1
                    Action := 51
                  Else 
                    Action := 52
                  Call Sub_AMR_MiR_V3
                  If AMR_Done
                    PROCESS_Step := 0
              Case (caseValue=2)
                Folder prepare
                  'THINGS THAT HAVE TO BE DONE ONCE IN A SEQUENCE,WORKFLOW'
                  PROCESS_Info := "prepare for work"
                  Script: log_process(PROCESS_Info)
                  If TASK.WORK.ITM_ID_Src>1
                    ITM_ID := TASK.WORK.ITM_ID_Src
                  ElseIf TASK.WORK.ITM_ID_Tgt>1
                    ITM_ID := TASK.WORK.ITM_ID_Tgt
                  If not ARM_Referenced and (ITM_ID≠0)
                    STP := 1
                  ElseIf ARM_Referenced or (ITM_ID≟0)
                    STP := 2
                  Switch expression=STP
                    Case (caseValue=1)
                      Folder reference [hidden by the author, left out]
                    Case (caseValue=2)
                      Folder manipulate [hidden by the author, left out]
                  ITM_Prepared := (ITM_Manipulated or  not found_in_list(ITM_ID, ITM_ID_List)) and (ARM_Referenced or ITM_ID≟0) and  not WRK_Done
                  STP := 0
                  STP_Info := ""
                  PROCESS_Step := 0
              Case (caseValue=3)
                Folder work
                  'ADD EVERY MACHINE, OBJECT, STATION TO WORK ON'
                  Switch expression=ITM_ID
                    Case (caseValue=1)
                      Folder uLM
                        If TASK.ID≟12
                          Folder fill racks
                            Action := 151
                            Call Sub_Vision_V18
                            If not ERROR.FLAG
                              Folder Actions for the task
                                Action := 1
                                JIG := 2
                                JIG_Slot := CAM_Result[0]
                                OBJ_Nbr := CAM_Result[0]
                                OBJ_Type := 2
                                Call Sub_Action_V4
                                If OBJ_Picked
                                  Script: CAM_Result.remove(0)
                                  PRC_TubCounter := PRC_TubCounter+1
                                  If PRC_TubCounter%4≟0
                                    JIG_Slot := 4
                                  Else 
                                    JIG_Slot := PRC_TubCounter%4
                                  OBJ_Nbr := ceil(PRC_TubCounter/4)
                                  Action := 2
                                  JIG := 4
                                  Call Sub_Action_V4
                                  Action := 151
                                  Call Sub_Vision_V18
                            If (CAM_Captures≥CAM_PRM_Retries) or (PRC_TubCounter≥32)
                              PROCESS_Step := 0
                              WRK_Done := True
                          SuppressedNode
                            Folder Transfering
                              Loop While (checkContinuously=false) expression=length(CAM_Result)>0 and CAM_Captures≤CAM_PRM_Retries and  not CMD_Stop and  not ERROR.FLAG
                                Placeholder
                        ElseIf TASK.ID≟10
                          Folder Pick Rack
                            Action := 131
                            Call Sub_Vision_V18
                            Action := 1
                            Call Sub_Action_V4
                            PROCESS_Step := 0
                            WRK_Done := True
                        ElseIf TASK.ID≟11
                          Folder Place Rack
                            Action := 2
                            Call Sub_Action_V4
                            PROCESS_Step := 0
                            WRK_Done := True
                        ElseIf TASK.ID≟13
                          Folder empty racks [hidden by the author, left out]
                        ElseIf TASK.ID≟14
                          SuppressedNode
                            Action := 131
                          SuppressedNode
                            Call Sub_Vision_V18
                          samples := True
                          Loop While (checkContinuously=false) expression=samples≟ True
                            SuppressedNode
                              JIG := 7
                            SuppressedNode
                              Action := 151
                            SuppressedNode
                              Call Sub_Vision_V18
                            SuppressedNode
                              Action := 1
                            SuppressedNode
                              Call Sub_Action_V4
                            JIG := 1
                            Action := 11
                            Call Sub_Action_V4
                            Action := 12
                            Call Sub_Action_V4
                            Action := 2
                            JIG := 6
                            Call Sub_Action_V4
                            Action := 13
                            Call Sub_Action_V4
                            Action := 1
                            JIG := 1
                            Call Sub_Action_V4
                            SuppressedNode
                              JIG := 7
                            SuppressedNode
                              Action := 2
                            SuppressedNode
                              Call Sub_Action_V4
                    Case (caseValue=2)
                      SuppressedNode
                        Folder Centrfiuge
                          SuppressedNode
                            Script: cent_error_check()
                          OBJ_Type := 1
                          If not ERROR.FLAG
                            'load racks'
                            If TASK.ID≟14
                              Loop While (checkContinuously=false) expression=(PRC_RackCounter<4) and  not CMD_Stop and  not ERROR.FLAG
                                ITM_ID := TASK.WORK.ITM_ID_Src
                                JIG := 4
                                JIG_Slot := PRC_RackCounter+1
                                Action := 1
                                Call Sub_Action_V4
                                If OBJ_Picked and  not ERROR.FLAG
                                  ITM_ID := TASK.WORK.ITM_ID_Tgt
                                  Script: execute_cent_action(ACTION_ROTATE, JIG_Slot)
                                  Action := 7
                                  Call Sub_Action_V4
                                  PRC_RackCounter := PRC_RackCounter + 1
                              If not ERROR.FLAG
                                WRK_Done := True
                                PROCESS_Step := 0
                            'unload racks'
                            If TASK.ID≟15
                              If CNT_State_Actual≟2 or CNT_State_Actual≟3
                                Loop While (checkContinuously=false) expression=(PRC_RackCounter<4) and  not CMD_Stop and  not ERROR.FLAG
                                  ITM_ID := TASK.WORK.ITM_ID_Src
                                  JIG_Slot := PRC_RackCounter + 1
                                  Script: execute_cent_action(ACTION_ROTATE, JIG_Slot)
                                  Script: execute_cent_action(ACTION_INSPECT, JIG_Slot)
                                  Action := 8
                                  Call Sub_Action_V4
                                  If OBJ_Picked and  not ERROR.FLAG
                                    ITM_ID := TASK.WORK.ITM_ID_Tgt
                                    JIG := 4
                                    JIG_Slot := PRC_RackCounter + 1
                                    Action := 2
                                    Call Sub_Action_V4
                                    PRC_RackCounter := PRC_RackCounter+1
                                If not ERROR.FLAG
                                  WRK_Done := True
                                  PROCESS_Step := 0
                    Case (caseValue=20)
                      SuppressedNode
                        Folder Biorad rack
                          'load racks'
                          If Task_ID≟16
                            SuppressedNode
                              PRC_RackCounter := 0
                            Loop While (checkContinuously=false) expression=(PRC_RackCounter<PRC_RackNumber) and  not CMD_Stop
                              JIG_Slot := PRC_RackCounter
                              Action := 1
                              PRC_Target := 0
                              Call Sub_Action_V4
                              If OBJ_Picked
                                Action := 2
                                PRC_Target := 1
                                Call Sub_Action_V4
                                Action := 7
                                PRC_Target := 1
                                Call Sub_Action_V4
                                PRC_RackCounter := PRC_RackCounter+1
                            WRK_Done := True
                            PROCESS_Step := 0
                          'unload racks'
                          SuppressedNode
                            If Task_ID≟17
                              SuppressedNode
                                PRC_RackCounter := 0
                              Loop While (checkContinuously=false) expression=(PRC_RackCounter<PRC_RackNumber) and  not CMD_Stop
                                JIG_Slot := PRC_RackCounter
                                Action := 8
                                PRC_Target := 1
                                Script: textmsg("Callactionunload=",Action)
                                Call Sub_Action_V4
                                Action := 1
                                PRC_Target := 1
                                Script: textmsg("Callactionpick=",Action)
                                Call Sub_Action_V4
                                If OBJ_Picked
                                  Action := 2
                                  PRC_Target := 0
                                  Script: textmsg("Callactionplace=",Action)
                                  Call Sub_Action_V4
                                  PRC_RackCounter := PRC_RackCounter+1
                              WRK_Done := True
                              PROCESS_Step := 0
                          If Task_ID≟17
                            PRC_RackCounter := 0
                            Loop While (checkContinuously=false) expression=(PRC_RackCounter<PRC_RackNumber) and  not CMD_Stop
                              Wait Condition expression=SensorData[PRC_RackCounter]≟1
                              JIG_Slot := PRC_RackCounter
                              Action := 8
                              PRC_Target := 1
                              Script: textmsg("Callactionunload=",Action)
                              Call Sub_Action_V4
                              Action := 1
                              PRC_Target := 1
                              Script: textmsg("Callactionpick=",Action)
                              Call Sub_Action_V4
                              If OBJ_Picked
                                Action := 2
                                PRC_Target := 0
                                Script: textmsg("Callactionplace=",Action)
                                Call Sub_Action_V4
                                PRC_RackCounter := PRC_RackCounter+1
                            WRK_Done := True
                            PROCESS_Step := 0
                    Case (caseValue=2147483647)
                      WRK_Done := True
                      PROCESS_Step := 0
          If CMD_Hold
            STATE := 9
            Script: ugo_update_outputs()
          ElseIf CMD_Suspend
            STATE := 12
            Script: ugo_update_outputs()
      Case (caseValue=7)
        Folder Completing [hidden by the author, left out]
      Case (caseValue=8)
        Folder Complete
          STATE_Info := "Complete"
          If CMD_Reset
            STATE := 3
            Script: ugo_update_outputs()
      Case (caseValue=9)
        Folder Holding [hidden by the author, left out]
      Case (caseValue=10)
        Folder Held [hidden by the author, left out]
      Case (caseValue=11)
        Folder Unholding [hidden by the author, left out]
      Case (caseValue=12)
        Folder Suspending [hidden by the author, left out]
      Case (caseValue=13)
        Folder Suspended [hidden by the author, left out]
      Case (caseValue=14)
        Folder Unsuspending [hidden by the author, left out]
      Case (caseValue=15)
        Folder Aborting [hidden by the author, left out]
      Case (caseValue=16)
        Folder Aborted [hidden by the author, left out]
      Case (caseValue=17)
        Folder Clearing [hidden by the author, left out]
    Script: log_state(STATE_Info)
    Script: log_warning(WARNING.MSG)
    Script: log_error(ERROR.MSG)
    Folder Times [hidden by the author, left out]
    SuppressedNode
      Script: sync()
    Wait Sleep waitTime=0.1
Thread Thread_1 (runOnlyOnce=false)
  BS_Error := GP_bool_in[10]
  SuppressedNode
    Set SingleDigitalPulseActionState SingleDigitalPulseActionState(hiPulseInSeconds=1, pin=GP_bool_out[1])
  BS_Busy := GP_bool_in[13]
  SuppressedNode
    If BS_Terminal≟ True
      Set DigitalOutput pin=digital_out[4]; digitalValue=1
      Set DigitalOutput pin=digital_out[2]; digitalValue=1
  BS_Complete := GP_bool_in[12]
  SuppressedNode
    If BS_Complete≟ True
      Set DigitalOutput pin=digital_out[4]; digitalValue=0
      Set DigitalOutput pin=digital_out[2]; digitalValue=0
      Set DigitalOutput pin=GP_bool_out[2]; digitalValue=1
  SuppressedNode
    Folder Folder
      SuppressedNode
        Set ExpressionOutput pin=GP_bool_out[0]; expression=digital_in[2]
      SuppressedNode
        Set ExpressionOutput pin=GP_bool_out[2]; expression=digital_in[3]
      SuppressedNode
        Wait Sleep waitTime=1
      SuppressedNode
        Set ExpressionOutput pin=GP_bool_out[2]; expression=False
      SuppressedNode
        Set ExpressionOutput pin=GP_bool_out[0]; expression=digital_in[2]
      SuppressedNode
        Set ExpressionOutput pin=GP_bool_out[1]; expression=digital_in[4]
  SuppressedNode
    Wait Sleep waitTime=4
  SuppressedNode
    Set DigitalOutput pin=GP_bool_out[2]; digitalValue=1
SubProgram -> Sub_Vision_V18
SubProgram  [hidden by the author, left out]
SubProgram -> Sub_Action_V4
SuppressedNode
  SubProgram Sub_Action_V1 (keepSynchronizedWithDisk=false) programFile=/programs/20241028 Robot Backup/03 Sub Routines/Sub_Action_V1.urp
    Folder PreSettings
      Folder init poses
        PSE_A := p[0,0,0,0,0,0]
        PSE_A_H := p[0,0,0,0,0,0]
        PSE_T := p[0,0,0,0,0,0]
        PSE_T_H := p[0,0,0,0,0,0]
        PSE_G := p[0,0,0,0,0,0]
        PSE_G_H := p[0,0,0,0,0,0]
        PSE_R := p[0,0,0,0,0,0]
        PSE_R_H := p[0,0,0,0,0,0]
        PSE_R_HH := p[0,0,0,0,0,0]
        PSE_R_HHH := p[0,0,0,0,0,0]
        JNT_A := [0,0,0,0,0,0]
        JNT_S := [0,0,0,0,0,0]
      PROCESS_Info := "work at target, Table"
      Folder Gripping parameters
        GRP_Open_Pose := 45
        GRP_Open_Pos_2 := 35
        GRP_Closed_Pose := 100
        Script: rq_set_force_norm(20)
        Script: rq_set_speed_norm(60)
      Switch expression=ITM_ID
        Case (caseValue=1)
          SuppressedNode
            Folder base plate uLM
              Script: FRM_Reference = ULM_Rack
              Folder Boxes [hidden by the author, left out]
          Folder uML
            Switch expression=JIG
              Case (caseValue=5)
                Folder 3finger gripper
                  Folder define poses
                    'Place in 3finger'
                    Script: FRM_Reference = ULM_3FG
                    PSE_T := pose_RPY2RotVec(p[0,0,0,0,0,0])
                    PSE_A := pose_trans(PSE_T, p[0,0,0.1,0,0,0])
                    PSE_R := pose_add(PSE_T, p[0,0,0.100,0,0,0])
                    If Action≟5
                      PSE_T := pose_RPY2RotVec(p[0,0,0.018,0,0,0])
                      PSE_T_H := pose_trans(PSE_T, p[0,0,0.02,0,0,0])
              Case (caseValue=6)
                Folder Caps bin
                  Folder define poses
                    'Drop cap'
                    Script: FRM_Reference=ULM_Bin
                    PSE_T := pose_RPY2RotVec(p[0,0,0,0,0,0])
                    PSE_T_H := pose_add(PSE_T, p[0,0,-0.011,0,0,0])
                    PSE_A := pose_trans(PSE_T, p[0,0,0.1,0,0,0])
                    PSE_R := pose_add(PSE_T, p[0,0,0.100,0,0,0])
              Case (caseValue=7)
                Folder define poses Manual
                  GRP_Open_Pose := 74
                  GRP_Open_Pos_2 := 74
                  FRM_Reference := ULM_Rack_tubes
                  PSE_T := pose_RPY2RotVec(p[0.0202*(JIG_Slot%10),0.0202*(floor(JIG_Slot/10)),0,0,0,0])
                  PSE_A := pose_trans(PSE_T, p[0,0,0.1,0,0,0])
                  PSE_R := pose_add(PSE_T, p[0,0,0.2500,0,0,0])
              Case (caseValue=8)
                Folder define poses Manual
                  GRP_Open_Pose := 74
                  GRP_Open_Pos_2 := 74
                  FRM_Reference := ULM_Rack_tubes
                  PSE_T := pose_RPY2RotVec(p[0.0202*(JIG_Slot%10),0.0202*(floor(JIG_Slot/10)),0,0,0,0])
                  PSE_A := pose_trans(PSE_T, p[0,0,0.1,0,0,0])
                  PSE_R := pose_add(PSE_T, p[0,0,0.100,0,0,0])
        Case (caseValue=2)
          SuppressedNode
            Folder pick area
              Switch expression=JIG
                Case (caseValue=1)
                  Folder Pick area for Atellica boxes
                    Script: FRM_Reference = FRM_PickUp_Atll
                    PSE_T := pose_RPY2RotVec(p[0.090,0.113,0.046,-40,0,90])
                Case (caseValue=2)
                  Folder Pick area for Atras boxes
                    Script: FRM_Reference = FRM_PickUp_Atrs
                    PSE_T := pose_RPY2RotVec(p[0.090,0.113,0.046,-40,0,90])
              Folder poses [hidden by the author, left out]
          Folder Sarstedt
            'CHANGE THE REFERENCE TO THE FRAME TO MOVE IN'
            Folder Gripping parameters
              GRP_Open_Pos := 45
              GRP_Close_Pos := 100
              Script: rq_set_force_norm(80)
              Script: rq_set_speed_norm(100)
            If PRC_Target≟0
              Script: FRM_Reference = ULM_Rack_Holder
              PSE_T := pose_RPY2RotVec(p[0,0,0,0,0,0])
              PSE_A := pose_trans(PSE_T, p[0,0,0.1,0,0,0])
              PSE_R := pose_add(PSE_T, p[0,0,0.1,0,0,0])
            Else 
              Script: FRM_Reference = FRM_DropOff
              PSE_T := pose_RPY2RotVec(p[0,0,0,0,0,0])
              PSE_A := pose_trans(PSE_T, p[0,0,0.1,0,0,0])
              PSE_R := pose_add(PSE_T, p[0,0,0.1,0,0,0])
      Folder Additional check
        If not is_reachable(FRM_Reference,[PSE_A,PSE_A_H,PSE_T,PSE_T_H,PSE_T_HH,PSE_R,PSE_R_H,PSE_R_HH,PSE_R_HHH])
          Folder Error [hidden by the author, left out]
          Action := 0
    Switch expression=Action
      Case (caseValue=1)
        Folder Pick [hidden by the author, left out]
      Case (caseValue=2)
        Folder Place [hidden by the author, left out]
      Case (caseValue=3)
        Folder Pick decapped probe from 3finger
          Action_Info := "Pick Rack/Probe"
          MoveJ speed 100 deg/s, acceleration 80 deg/s^2 (useActiveTCP=true) feature=FRM_Reference
            Waypoint Variable (Variable): variable=PSE_A
          Script: rq_move_and_wait_norm(GRP_Open_Pose)
          MoveL speed 75 mm/s, acceleration 150 mm/s^2 (useActiveTCP=true) feature=FRM_Reference
            SuppressedNode
              Script: PSE_T[2]=PSE_T[2]-0.005
            Waypoint Variable (Variable): variable=PSE_T
            SuppressedNode
              Force Frame feature=FRM_Reference; selection=[1, 1, 0, 0, 0, 0]; wrench=[0, 0, 0, 0, 0, 0]; limitsForce=[0.25, 0.25, 0.15, 1.047198, 1.047198, 1.047198]; limitsMotion=[0.1, 0.1, 0.1, 0.349066, 0.349066, 0.349066]
                Waypoint Variable (Variable): motionParameters(jointSpeed=1.047198 jointAcceleration=1.396263 cartesianSpeed=0.03 cartesianAcceleration=0.2); variable=PSE_T
            'ADD OPEN GRIPPER'
            Script: rq_set_force_norm(20)
            Script: rq_set_speed_norm(30)
            Script: rq_move_and_wait_norm(GRP_Closed_Pose)
          Set DigitalOutput pin=digital_out[5]; digitalValue=1
          Wait Sleep waitTime=0.3
          MoveL speed 100 mm/s, acceleration 1200 mm/s^2 (useActiveTCP=true) feature=FRM_Reference
            Waypoint Variable (Variable): motionParameters(jointSpeed=1.047198 jointAcceleration=1.396263 cartesianSpeed=0.25 cartesianAcceleration=1.2); variable=PSE_R
      Case (caseValue=4)
        Folder Place probe in 3finger
          Action_Info := "place object"
          MoveJ speed 100 deg/s, acceleration 80 deg/s^2 (useActiveTCP=true) feature=FRM_Reference
            Waypoint Variable (Variable): variable=PSE_A
          Set DigitalOutput pin=digital_out[5]; digitalValue=1
          MoveL speed 75 mm/s, acceleration 150 mm/s^2 (useActiveTCP=true) feature=FRM_Reference
            Waypoint Variable (Variable): variable=PSE_T
              Until TOOL_CONTACT_DETECTION (allowActions=false retraction=0 decelerationAcceleration=3 decelerationAngularAcceleration=34.906585)
          Set DigitalOutput pin=digital_out[5]; digitalValue=0
          Wait Sleep waitTime=0.15
          SuppressedNode
            If Task_ID≟12
              Wait Sleep waitTime=0.15
              MoveL speed 75 mm/s, acceleration 150 mm/s^2 (useActiveTCP=true) feature=FRM_Reference
                Waypoint Variable (Variable): variable=PSE_R
      Case (caseValue=5)
        SuppressedNode
          Folder Decapping
            Action_Info := "decapping"
            PRC_decap_z_val := z_Pos
            PRM_forcdistSta := 0.024
            Script: zero_ftsensor()
            Wait Sleep waitTime=1
            Set DigitalOutput pin=EN_3FG_Motor; digitalValue=1
            Set DigitalOutput pin=Decap_3FG; digitalValue=1
            Force Frame feature=ULM_3FG; selection=[0, 0, 1, 0, 0, 0]; wrench=[0, 0, 20, 0, 0, 0]; limitsForce=[0.04, 0.04, 0.015, 1.047198, 1.047198, 1.047198]; limitsMotion=[0.1, 0.1, 0.1, 0.349066, 0.349066, 0.349066]
              PRC_Force := True
              Wait Condition expression=PRM_forcdistLiv>PRM_forcdistSta
            PRC_Force := False
            Set DigitalOutput pin=EN_3FG_Motor; digitalValue=0
            Set DigitalOutput pin=Decap_3FG; digitalValue=0
            MoveL speed 150 mm/s, acceleration 800 mm/s^2 (useActiveTCP=true) feature=FRM_Reference
              Waypoint Variable (Variable): variable=PSE_R
      Case (caseValue=6)
        Folder Drop the cap
          If JNT_A≠[0,0,0,0,0,0]
            MoveJ speed 100 deg/s, acceleration 80 deg/s^2 (useActiveTCP=true positionType=JointAngles) feature=FRM_Reference
              Waypoint Variable (Variable): motionParameters(blendRadius=0.02); variable=JNT_A
          Else 
            MoveJ speed 100 deg/s, acceleration 80 deg/s^2 (useActiveTCP=true) feature=FRM_Reference
              Waypoint Variable (Variable): motionParameters(blendRadius=0.02); variable=PSE_A
          MoveL speed 400 mm/s, acceleration 500 mm/s^2 (useActiveTCP=true) feature=FRM_Reference
            Waypoint Variable (Variable): motionParameters(jointSpeed=1.047198 jointAcceleration=1.396263 cartesianSpeed=0.09 cartesianAcceleration=0.05); variable=PSE_T
            'ADD OPEN GRIPPER'
            URCap Gripper (Robotiq_Grippers, Robotiq Inc.) dataModel(position=78.82352941176471, force=11.0, speed=0.0, positionInDouble=78.82352941176471, forceInDouble=11.0, speedInDouble=0.0, slaveIds=[9], blocking=true)
            Waypoint Variable (Variable): motionParameters(jointSpeed=1.047198 jointAcceleration=1.396263 cartesianSpeed=0.09 cartesianAcceleration=0.05); variable=PSE_T_H
            URCap Gripper (Robotiq_Grippers, Robotiq Inc.) dataModel(position=24.705882352941178, force=11.0, speed=0.0, positionInDouble=24.705882352941178, forceInDouble=11.0, speedInDouble=0.0, slaveIds=[9], blocking=true)
            SuppressedNode
              URCap Gripper (Robotiq_Grippers, Robotiq Inc.) dataModel(position=100.0, force=28.0, speed=100.0, positionInDouble=100.0, forceInDouble=28.0, speedInDouble=100.0, slaveIds=[9], blocking=true)
            SuppressedNode
              Wait Sleep waitTime=0.2
            SuppressedNode
              Loop While (checkContinuously=false) expression=rq_is_object_detected()
                Script: rq_set_force_norm(10)
                Script: rq_set_speed_norm(100)
                URCap Gripper (Robotiq_Grippers, Robotiq Inc.) dataModel(position=0.0, force=28.0, speed=100.0, positionInDouble=0.0, forceInDouble=28.0, speedInDouble=100.0, slaveIds=[9], blocking=true)
                Wait Sleep waitTime=0.5
                URCap Gripper (Robotiq_Grippers, Robotiq Inc.) dataModel(position=100.0, force=28.0, speed=100.0, positionInDouble=100.0, forceInDouble=28.0, speedInDouble=100.0, slaveIds=[9], blocking=true)
            SuppressedNode
              Wait Sleep waitTime=0.2
            Waypoint Variable (Variable): variable=PSE_R
      Case (caseValue=16)
        Folder Scan the barcode
          Action_Info := "scan the barcode"
          Barc_scan_succs := False
          Folder First check
            Set DigitalOutput pin=GP_bool_out[1]; digitalValue=1
            Wait Sleep waitTime=0.1
            Barc_scan_succs := digital_in[6]
          If Barc_scan_succs
            Set DigitalOutput pin=digital_out[5]; digitalValue=1
            Set DigitalOutput pin=digital_out[2]; digitalValue=1
            Loop While (checkContinuously=true) expression=Barc_scan_succs
              Barc_scan_succs := digital_in[6]
              Wait Sleep waitTime=0.05
            Set DigitalOutput pin=digital_out[5]; digitalValue=0
            Set DigitalOutput pin=digital_out[2]; digitalValue=0
            Set DigitalOutput pin=digital_out[6]; digitalValue=0
          Else 
            Timer (action=Reset) variable(name=Timer_Barc_scan)
            Timer (action=Start) variable=Timer_Barc_scan
            Set DigitalOutput pin=digital_out[3]; digitalValue=1
            Set DigitalOutput pin=digital_out[5]; digitalValue=1
            Loop While (checkContinuously=true) expression=not Barc_scan_succs and  not CMD_Stop and Timer_Barc_scan<60
              SuppressedNode
                If Timer_Barc_scan>1.5
                  Placeholder
              Set DigitalOutput pin=digital_out[6]; digitalValue=1
              Barc_scan_succs := digital_in[6]
              Wait Sleep waitTime=0.05
            Set DigitalOutput pin=digital_out[5]; digitalValue=0
            Set DigitalOutput pin=digital_out[3]; digitalValue=0
            Set DigitalOutput pin=digital_out[6]; digitalValue=0
            Timer (action=Stop) variable=Timer_Barc_scan
            If Timer_Barc_scan≥60
              Script: set_error(5200)
    '=========='
    Folder PostSettings [hidden by the author, left out]
SuppressedNode
  SubProgram Sub_Action_V2 (keepSynchronizedWithDisk=false) programFile=/programs/03 Sub Routines/SubAction_V2/Sub_Action_V2.urp
    Folder PreSettings
      Folder init poses
        PSE_A := p[0,0,0,0,0,0]
        PSE_A_H := p[0,0,0,0,0,0]
        PSE_T := p[0,0,0,0,0,0]
        PSE_T_H := p[0,0,0,0,0,0]
        PSE_G := p[0,0,0,0,0,0]
        PSE_G_H := p[0,0,0,0,0,0]
        PSE_R := p[0,0,0,0,0,0]
        PSE_R_H := p[0,0,0,0,0,0]
        JNT_A := [0,0,0,0,0,0]
        JNT_S := [0,0,0,0,0,0]
        JNT_Q := [0,0,0,0,0,0]
      PROCESS_Info := "work at target, Table"
      PRM_TubHghtDiff := -0.024
      Folder Gripping parameters
        GRP_Open_Pos := 45
        GRP_Close_Pos := 100
        Script: rq_set_force_norm(20)
        Script: rq_set_speed_norm(80)
      Switch expression=ITM_ID
        Case (caseValue=1)
          Folder uML
            Switch expression=JIG
              Case (caseValue=2)
                Folder biorad rack tubes
                  GRP_Open_Pos := 60
                  FRM_Reference := uLM_BradRckTubs
                  Tubes_in_Rack := 6
                  PSE_T := pose_RPY2RotVec(p[0.02*(JIG_Slot%Tubes_in_Rack),-0.04365*floor(JIG_Slot/Tubes_in_Rack),0.003,0,0,-90])
                  SuppressedNode
                    Script: PSE_T[2]=PSE_T[2]+PRM_TubHghtDiff
                  If (JIG_Slot%Tubes_in_Rack)>1
                    Script: PSE_T[0]=PSE_T[0]+0.0165
                    If (JIG_Slot%Tubes_in_Rack)>4
                      Script: PSE_T[0]=PSE_T[0]+0.0235
                      SuppressedNode
                        If (JIG_Slot%10)>6
                          Script: PSE_T[0]=PSE_T[0]+0.0165
                  PSE_R := pose_add(PSE_T, p[0,0,0.2500,0,0,0])
                  PSE_A := pose_add(PSE_T, p[0,0,0.1,0,0,0])
              Case (caseValue=4)
                Folder centrifuge rack tubes
                  GRP_Open_Pos := 60
                  FRM_Reference := uLM_CentTubes
                  PSE_T := pose_RPY2RotVec(p[0.0975*(JIG_Slot%4),0,0.002,0,0,0])
                  SuppressedNode
                    Script: PSE_T[2]=PSE_T[2]+PRM_TubHghtDiff
                  If JIG_Slot>3 and JIG_Slot≤7
                    Script: PSE_T[1]=0.06
                    Script: PSE_T[0]=PSE_T[0]+0.06
                  ElseIf JIG_Slot>7 and JIG_Slot≤11
                    Script: PSE_T[0]=PSE_T[0]+0.06
                  ElseIf JIG_Slot>11 and JIG_Slot≤15
                    Script: PSE_T[1]=0.06
                  PSE_R := pose_add(PSE_T, p[0,0,0.150,0,0,0])
                  PSE_A := pose_add(PSE_T, p[0,0,0.15,0,0,0])
                  JNT_Q := [-1.4,-1.89,-1.4,-1.42,1.57,0.18]
              Case (caseValue=5)
                Folder 3finger gripper
                  Folder define poses
                    'Place in 3finger'
                    Script: FRM_Reference = uML_3fingergrip
                    PSE_T := pose_RPY2RotVec(p[0,0,0.003,0,0,0])
                    Script: PSE_T[2]=PSE_T[2]+PRM_TubHghtDiff
                    If Action≟5
                      PSE_T := pose_RPY2RotVec(p[0,0,0.018,0,0,0])
                      PSE_T_H := pose_trans(PSE_T, p[0,0,0.02,0,0,0])
                    If Action≟3
                      Script: PSE_T[5]=PSE_T[5]+d2r(155)
                    PSE_A := pose_trans(PSE_T, p[0,0,0.1,0,0,0])
                    PSE_R := pose_add(PSE_T, p[0,0,0.060,0,0,0])
              Case (caseValue=6)
                Folder Caps bin
                  Folder define poses
                    'Drop cap'
                    Script: FRM_Reference=uML_CapBin
                    SuppressedNode
                      PSE_T := pose_RPY2RotVec(p[0.037,0,0.005,0,0,0])
                    PSE_T := pose_RPY2RotVec(p[0,0,0.005,0,0,0])
                    PSE_T_H := pose_trans(PSE_T, p[0,0,-0.008,0,0,0])
                    PSE_A := pose_trans(PSE_T, p[0,0,0.1,0,0,0])
                    PSE_R := pose_add(PSE_T, p[0,0,0.100,0,0,0])
              Case (caseValue=7)
                Folder define poses Manual
                  GRP_Open_Pos := 60
                  FRM_Reference := uLM_Manual
                  If Action≟1
                    SuppressedNode
                      PSE_T := pose_RPY2RotVec(p[0.0202*(JIG_Slot%10),0.0202*(floor(JIG_Slot/10)),0,0,0,0])
                    PSE_T := pose_RPY2RotVec(p[0.0248*(JIG_Slot%8),0.0258*(floor(JIG_Slot/8)),0,0,0,0])
                    PSE_R := pose_add(PSE_T, p[0,0,0.150,0,0,0])
                  ElseIf Action≟2
                    SuppressedNode
                      PSE_T := pose_RPY2RotVec(p[0.0202*(JIG_Slot%10),0.0202*(floor(JIG_Slot/10)),0,0,0,-62])
                    PSE_T := pose_RPY2RotVec(p[0.0248*(JIG_Slot%8),0.0258*(floor(JIG_Slot/8)),0,0,0,0])
                    PSE_R := pose_add(PSE_T, p[0,0,0.100,0,0,0])
                  Script: PSE_T[2]=PSE_T[2]+PRM_TubHghtDiff
                  PSE_A := pose_add(PSE_T, p[0,0,0.1,0,0,0])
        Case (caseValue=2)
          Folder Biorad
            'CHANGE THE REFERENCE TO THE FRAME TO MOVE IN'
            Folder Gripping parameters [hidden by the author, left out]
            If PRC_Target≟0
              Script: FRM_Reference = uML_BradRacks
              PSE_T := pose_RPY2RotVec(p[0.04365*JIG_Slot,0,0,0,0,180])
              If Action≟2
                SuppressedNode
                  Script: PSE_T[2]=PSE_T[2]+0.008
                Script: PSE_T[2]=PSE_T[2]+0.002
              PSE_A := pose_add(PSE_T, p[0,0,0.18,0,0,0])
              PSE_R := pose_add(PSE_T, p[0,0,0.18,0,0,0])
            Else 
              Script: FRM_Reference = FRM_BioradMachn
              Switch expression=Action
                Case (caseValue=1)
                  PSE_T := pose_RPY2RotVec(p[0.125-0.056*JIG_Slot,0.07,0.139,-90,0,0])
                  PSE_A := pose_add(PSE_T, p[0,0.1,0,0,0,0])
                  PSE_R := pose_add(PSE_T, p[0,0.05,0.1,0,0,0])
                Case (caseValue=2)
                  PSE_T := pose_RPY2RotVec(p[0.125-0.056*JIG_Slot,0.07,0.08,-90,0,0])
                  PSE_T_H := pose_RPY2RotVec(p[0.125-0.056*JIG_Slot,0.072,0.238,-90,0,0])
                  PSE_A := pose_add(PSE_T_H, p[0,0.1,0,0,0,0])
                  PSE_R := pose_add(PSE_T_H, p[0,0.1,0,0,0,0])
                Case (caseValue=7)
                  PSE_T := pose_RPY2RotVec(p[0.124-0.056*JIG_Slot,0.084,0.008,-55,0,0])
                  PSE_T_H := pose_RPY2RotVec(p[0.125-0.056*JIG_Slot,0.084,0.284,-55,0,0])
                  PSE_A := pose_add(PSE_T_H, p[0,0.05,0.05,0,0,0])
                  PSE_R := pose_add(PSE_T, p[0,0,0.1,0,0,0])
                  SuppressedNode
                    JNT_Q := [0.108,-1.505,-1.993,-0.886,1.488,3.189]
                Case (caseValue=8)
                  PSE_T_H := pose_RPY2RotVec(p[0.124-0.056*JIG_Slot,0.092,0.049,-72,0,0])
                  PSE_T := pose_RPY2RotVec(p[0.125-0.056*JIG_Slot,0.092,0.316,-72,0,0])
                  PSE_R := pose_add(PSE_T, p[0,0.05,0,0,0,0])
                  PSE_A := pose_add(PSE_T_H, p[0,0,0.1,0,0,0])
                  JNT_Q := [0.108,-1.505,-1.993,-0.886,1.488,3.189]
                  If JIG_Slot≟0
                    Script: PSE_T[0]=PSE_T[0]-0.002
                    Script: PSE_T_H[0]=PSE_T_H[0]-0.002
        Case (caseValue=4)
          Folder Centrifuge
            'CHANGE THE REFERENCE TO THE FRAME TO MOVE IN'
            Folder Gripping parameters [hidden by the author, left out]
            If PRC_Target≟0
              Script: FRM_Reference = uLM_CentRacks
              Switch expression=Action
                Case (caseValue=1)
                  PSE_T := pose_RPY2RotVec(p[0.0975*(JIG_Slot%4),0,-0.015,0,0,0])
                Case (caseValue=2)
                  PSE_T := pose_RPY2RotVec(p[0.0975*(JIG_Slot%4),0,0.01,0,0,0])
              PSE_A := pose_add(PSE_T, p[0,0,0.15,0,0,0])
              PSE_R := pose_add(PSE_T, p[0,0,0.15,0,0,0])
            Else 
              Script: FRM_Reference = FRM_Centrifuge
              Switch expression=Action
                Case (caseValue=1)
                  PSE_T := pose_RPY2RotVec(p[0,0,-0.02,0,0,0])
                Case (caseValue=2)
                  PSE_T := pose_RPY2RotVec(p[0,0,0.015,0,0,0])
              PSE_A := pose_add(PSE_T, p[0,0,0.2,0,0,0])
              PSE_R := pose_add(PSE_T, p[0,0,0.25,0,0,0])
      Folder Additional check
        If not is_reachable(FRM_Reference,[PSE_A,PSE_A_H,PSE_T,PSE_T_H,PSE_R,PSE_R_H])
          Script: set_error(1002)
          Action := 0
    Switch expression=Action
      Case (caseValue=1)
        Folder Pick
          Action_Info := "Pick Rack/Probe"
          Script: do_transition(pose_trans(FRM_Reference, PSE_T), keep_rxry=OBJ_Picked)
          If not OBJ_Picked
            Script: rq_move_and_wait_norm(GRP_Open_Pos)
          If JNT_Q≠JNT_Z
            Script: movej(get_inverse_kin(pose_trans(FRM_Reference, PSE_A), qnear=JNT_Q))
          Else 
            MoveJ speed 100 deg/s, acceleration 80 deg/s^2 (useActiveTCP=true) feature=FRM_Reference
              Waypoint Variable (Variable): variable=PSE_A
          If ITM_ID≟4 and PRC_Target≟1
            Script: execute_cent_action(eACT_Inspect,(JIG_Slot+1))
          MoveL speed 400 mm/s, acceleration 500 mm/s^2 (useActiveTCP=true) feature=FRM_Reference
            Waypoint Variable (Variable): motionParameters(jointSpeed=1.047198 jointAcceleration=1.396263 cartesianSpeed=0.12 cartesianAcceleration=0.08); variable=PSE_T
            Script: rq_set_force_norm(50)
            SuppressedNode
              Script: rq_move_and_wait_norm(GRP_Close_Pos)
            URCap Gripper (Robotiq_Grippers, Robotiq Inc.) dataModel(position=100.0, force=76.0, speed=100.0, positionInDouble=100.0, forceInDouble=76.0, speedInDouble=100.0, slaveIds=[9], blocking=true)
            OBJ_Picked := rq_is_object_detected()
            Script: textmsg("Obj_Picked=",OBJ_Picked)
            If OBJ_Picked
              If PSE_T_H≠PSE_Z
                Waypoint Variable (Variable): motionParameters(blendRadius=0.01); variable=PSE_T_H
              Waypoint Variable (Variable): variable=PSE_R
            Else 
              Script: set_error(1010)
      Case (caseValue=2)
        Folder Place
          Action_Info := "place object"
          SuppressedNode
            Script: do_transition(keep_rxry=OBJ_Picked)
          Script: do_transition(pose_trans(FRM_Reference, PSE_T), keep_rxry=OBJ_Picked)
          If JNT_A≠[0,0,0,0,0,0]
            MoveJ speed 100 deg/s, acceleration 80 deg/s^2 (useActiveTCP=true positionType=JointAngles) feature=FRM_Reference
              Waypoint Variable (Variable): motionParameters(blendRadius=0.02); variable=JNT_A
          Else 
            MoveJ speed 100 deg/s, acceleration 80 deg/s^2 (useActiveTCP=true) feature=FRM_Reference
              Waypoint Variable (Variable): variable=PSE_A
          MoveL speed 400 mm/s, acceleration 500 mm/s^2 (useActiveTCP=true) feature=FRM_Reference
            If PSE_T_H≠PSE_Z
              Waypoint Variable (Variable): motionParameters(jointSpeed=1.047198 jointAcceleration=1.396263 cartesianSpeed=0.07 cartesianAcceleration=0.04); variable=PSE_T_H
            If ITM_ID≟4 and PRC_Target≟1
              Script: execute_cent_action(eACT_Inspect,(JIG_Slot+1))
            If not ERROR.FLAG
              If (ITM_ID≟1 and (JIG≟4 or JIG≟2)) or ITM_ID≟2 or ITM_ID≟4
                Waypoint Variable (Variable): motionParameters(jointSpeed=1.047198 jointAcceleration=1.396263 cartesianSpeed=0.09 cartesianAcceleration=0.05); variable=PSE_T
              Else 
                Waypoint Variable (Variable): motionParameters(jointSpeed=1.047198 jointAcceleration=1.396263 cartesianSpeed=0.09 cartesianAcceleration=0.05); variable=PSE_T
                  Until TOOL_CONTACT_DETECTION (allowActions=false retraction=0 decelerationAcceleration=0.5 decelerationAngularAcceleration=34.906585)
                Force Frame feature=FRM_Reference; selection=[1, 1, 0, 0, 0, 0]; wrench=[0, 0, 0, 0, 0, 0]; limitsForce=[0.05, 0.05, 0.15, 1.047198, 1.047198, 1.047198]; limitsMotion=[0.1, 0.1, 0.1, 0.349066, 0.349066, 0.349066]
                  Waypoint Variable (Variable): motionParameters(jointSpeed=1.047198 jointAcceleration=1.396263 cartesianSpeed=0.07 cartesianAcceleration=0.04); variable=PSE_T
              Script: rq_move_and_wait_norm(GRP_Open_Pos)
              Wait Sleep waitTime=0.2
              Waypoint Variable (Variable): variable=PSE_R
          SuppressedNode
            PRC_Task_Boxes := PRC_Task_Boxes+GRP_Boxes_Numb
      Case (caseValue=3)
        Folder Pick decapped probe from 3finger
          Action_Info := "Pick Rack/Probe"
          MoveJ speed 100 deg/s, acceleration 80 deg/s^2 (useActiveTCP=true) feature=FRM_Reference
            Waypoint Variable (Variable): variable=PSE_A
          Script: rq_move_and_wait_norm(GRP_Open_Pos)
